(* IEC 61131-3 sources: STAR-PLC-Agent/results/raw/codex_matrix_resume_20261114/codex_deepseek/SELF011/functional/attempt_0001, 1 file *)

(* ---- test_program.st ---- *)
PROGRAM PLC_PRG
VAR
 BenchStep : UDINT := 0;
 BenchCalls : UDINT := 0;
 BenchDone : BOOL := FALSE;
 BenchUut0 : FB_Task;
 BenchUut1 : FB_Task;
 BenchUut2 : FB_Task;
 BenchUut3 : FB_Task;
 BenchUut4 : FB_Task;
 BenchUut5 : FB_Task;
 BenchUut6 : FB_Task;
 BenchUut7 : FB_Task;
 BenchUut8 : FB_Task;
 BenchUut9 : FB_Task;
 BenchUut10 : FB_Task;
 BenchUut11 : FB_Task;
 TraceIn_Start : ARRAY[0..147] OF BOOL;
 TraceIn_Stop : ARRAY[0..147] OF BOOL;
 TraceIn_Reset : ARRAY[0..147] OF BOOL;
 TraceIn_ExtendDone : ARRAY[0..147] OF BOOL;
 TraceIn_ClampDone : ARRAY[0..147] OF BOOL;
 TraceIn_ReleaseDone : ARRAY[0..147] OF BOOL;
 TraceIn_RetractDone : ARRAY[0..147] OF BOOL;
 TraceOut_Extend : ARRAY[0..147] OF BOOL;
 TraceOut_Clamp : ARRAY[0..147] OF BOOL;
 TraceOut_Release : ARRAY[0..147] OF BOOL;
 TraceOut_Retract : ARRAY[0..147] OF BOOL;
 TraceOut_Busy : ARRAY[0..147] OF BOOL;
 TraceOut_Done : ARRAY[0..147] OF BOOL;
END_VAR

IF NOT BenchDone THEN
 CASE BenchStep OF
 0:
   BenchUut0.Start := TRUE;
   BenchUut0.Stop := FALSE;
   BenchUut0.Reset := FALSE;
   BenchUut0.ExtendDone := FALSE;
   BenchUut0.ClampDone := FALSE;
   BenchUut0.ReleaseDone := FALSE;
   BenchUut0.RetractDone := FALSE;
   TraceIn_Start[0] := BenchUut0.Start;
   TraceIn_Stop[0] := BenchUut0.Stop;
   TraceIn_Reset[0] := BenchUut0.Reset;
   TraceIn_ExtendDone[0] := BenchUut0.ExtendDone;
   TraceIn_ClampDone[0] := BenchUut0.ClampDone;
   TraceIn_ReleaseDone[0] := BenchUut0.ReleaseDone;
   TraceIn_RetractDone[0] := BenchUut0.RetractDone;
   BenchUut0();
   TraceOut_Extend[0] := BenchUut0.Extend;
   TraceOut_Clamp[0] := BenchUut0.Clamp;
   TraceOut_Release[0] := BenchUut0.Release;
   TraceOut_Retract[0] := BenchUut0.Retract;
   TraceOut_Busy[0] := BenchUut0.Busy;
   TraceOut_Done[0] := BenchUut0.Done;
   BenchCalls := BenchCalls + 1;
 1:
   BenchUut0.Start := TRUE;
   BenchUut0.Stop := FALSE;
   BenchUut0.Reset := FALSE;
   BenchUut0.ExtendDone := FALSE;
   BenchUut0.ClampDone := FALSE;
   BenchUut0.ReleaseDone := FALSE;
   BenchUut0.RetractDone := TRUE;
   TraceIn_Start[1] := BenchUut0.Start;
   TraceIn_Stop[1] := BenchUut0.Stop;
   TraceIn_Reset[1] := BenchUut0.Reset;
   TraceIn_ExtendDone[1] := BenchUut0.ExtendDone;
   TraceIn_ClampDone[1] := BenchUut0.ClampDone;
   TraceIn_ReleaseDone[1] := BenchUut0.ReleaseDone;
   TraceIn_RetractDone[1] := BenchUut0.RetractDone;
   BenchUut0();
   TraceOut_Extend[1] := BenchUut0.Extend;
   TraceOut_Clamp[1] := BenchUut0.Clamp;
   TraceOut_Release[1] := BenchUut0.Release;
   TraceOut_Retract[1] := BenchUut0.Retract;
   TraceOut_Busy[1] := BenchUut0.Busy;
   TraceOut_Done[1] := BenchUut0.Done;
   BenchCalls := BenchCalls + 1;
 2:
   BenchUut0.Start := FALSE;
   BenchUut0.Stop := FALSE;
   BenchUut0.Reset := FALSE;
   BenchUut0.ExtendDone := FALSE;
   BenchUut0.ClampDone := FALSE;
   BenchUut0.ReleaseDone := FALSE;
   BenchUut0.RetractDone := FALSE;
   TraceIn_Start[2] := BenchUut0.Start;
   TraceIn_Stop[2] := BenchUut0.Stop;
   TraceIn_Reset[2] := BenchUut0.Reset;
   TraceIn_ExtendDone[2] := BenchUut0.ExtendDone;
   TraceIn_ClampDone[2] := BenchUut0.ClampDone;
   TraceIn_ReleaseDone[2] := BenchUut0.ReleaseDone;
   TraceIn_RetractDone[2] := BenchUut0.RetractDone;
   BenchUut0();
   TraceOut_Extend[2] := BenchUut0.Extend;
   TraceOut_Clamp[2] := BenchUut0.Clamp;
   TraceOut_Release[2] := BenchUut0.Release;
   TraceOut_Retract[2] := BenchUut0.Retract;
   TraceOut_Busy[2] := BenchUut0.Busy;
   TraceOut_Done[2] := BenchUut0.Done;
   BenchCalls := BenchCalls + 1;
 3:
   BenchUut0.Start := FALSE;
   BenchUut0.Stop := FALSE;
   BenchUut0.Reset := FALSE;
   BenchUut0.ExtendDone := TRUE;
   BenchUut0.ClampDone := FALSE;
   BenchUut0.ReleaseDone := FALSE;
   BenchUut0.RetractDone := FALSE;
   TraceIn_Start[3] := BenchUut0.Start;
   TraceIn_Stop[3] := BenchUut0.Stop;
   TraceIn_Reset[3] := BenchUut0.Reset;
   TraceIn_ExtendDone[3] := BenchUut0.ExtendDone;
   TraceIn_ClampDone[3] := BenchUut0.ClampDone;
   TraceIn_ReleaseDone[3] := BenchUut0.ReleaseDone;
   TraceIn_RetractDone[3] := BenchUut0.RetractDone;
   BenchUut0();
   TraceOut_Extend[3] := BenchUut0.Extend;
   TraceOut_Clamp[3] := BenchUut0.Clamp;
   TraceOut_Release[3] := BenchUut0.Release;
   TraceOut_Retract[3] := BenchUut0.Retract;
   TraceOut_Busy[3] := BenchUut0.Busy;
   TraceOut_Done[3] := BenchUut0.Done;
   BenchCalls := BenchCalls + 1;
 4:
   BenchUut0.Start := FALSE;
   BenchUut0.Stop := FALSE;
   BenchUut0.Reset := FALSE;
   BenchUut0.ExtendDone := FALSE;
   BenchUut0.ClampDone := TRUE;
   BenchUut0.ReleaseDone := FALSE;
   BenchUut0.RetractDone := FALSE;
   TraceIn_Start[4] := BenchUut0.Start;
   TraceIn_Stop[4] := BenchUut0.Stop;
   TraceIn_Reset[4] := BenchUut0.Reset;
   TraceIn_ExtendDone[4] := BenchUut0.ExtendDone;
   TraceIn_ClampDone[4] := BenchUut0.ClampDone;
   TraceIn_ReleaseDone[4] := BenchUut0.ReleaseDone;
   TraceIn_RetractDone[4] := BenchUut0.RetractDone;
   BenchUut0();
   TraceOut_Extend[4] := BenchUut0.Extend;
   TraceOut_Clamp[4] := BenchUut0.Clamp;
   TraceOut_Release[4] := BenchUut0.Release;
   TraceOut_Retract[4] := BenchUut0.Retract;
   TraceOut_Busy[4] := BenchUut0.Busy;
   TraceOut_Done[4] := BenchUut0.Done;
   BenchCalls := BenchCalls + 1;
 5:
   BenchUut0.Start := FALSE;
   BenchUut0.Stop := FALSE;
   BenchUut0.Reset := FALSE;
   BenchUut0.ExtendDone := FALSE;
   BenchUut0.ClampDone := FALSE;
   BenchUut0.ReleaseDone := TRUE;
   BenchUut0.RetractDone := FALSE;
   TraceIn_Start[5] := BenchUut0.Start;
   TraceIn_Stop[5] := BenchUut0.Stop;
   TraceIn_Reset[5] := BenchUut0.Reset;
   TraceIn_ExtendDone[5] := BenchUut0.ExtendDone;
   TraceIn_ClampDone[5] := BenchUut0.ClampDone;
   TraceIn_ReleaseDone[5] := BenchUut0.ReleaseDone;
   TraceIn_RetractDone[5] := BenchUut0.RetractDone;
   BenchUut0();
   TraceOut_Extend[5] := BenchUut0.Extend;
   TraceOut_Clamp[5] := BenchUut0.Clamp;
   TraceOut_Release[5] := BenchUut0.Release;
   TraceOut_Retract[5] := BenchUut0.Retract;
   TraceOut_Busy[5] := BenchUut0.Busy;
   TraceOut_Done[5] := BenchUut0.Done;
   BenchCalls := BenchCalls + 1;
 6:
   BenchUut0.Start := FALSE;
   BenchUut0.Stop := FALSE;
   BenchUut0.Reset := FALSE;
   BenchUut0.ExtendDone := FALSE;
   BenchUut0.ClampDone := FALSE;
   BenchUut0.ReleaseDone := FALSE;
   BenchUut0.RetractDone := TRUE;
   TraceIn_Start[6] := BenchUut0.Start;
   TraceIn_Stop[6] := BenchUut0.Stop;
   TraceIn_Reset[6] := BenchUut0.Reset;
   TraceIn_ExtendDone[6] := BenchUut0.ExtendDone;
   TraceIn_ClampDone[6] := BenchUut0.ClampDone;
   TraceIn_ReleaseDone[6] := BenchUut0.ReleaseDone;
   TraceIn_RetractDone[6] := BenchUut0.RetractDone;
   BenchUut0();
   TraceOut_Extend[6] := BenchUut0.Extend;
   TraceOut_Clamp[6] := BenchUut0.Clamp;
   TraceOut_Release[6] := BenchUut0.Release;
   TraceOut_Retract[6] := BenchUut0.Retract;
   TraceOut_Busy[6] := BenchUut0.Busy;
   TraceOut_Done[6] := BenchUut0.Done;
   BenchCalls := BenchCalls + 1;
 7:
   BenchUut0.Start := TRUE;
   BenchUut0.Stop := FALSE;
   BenchUut0.Reset := FALSE;
   BenchUut0.ExtendDone := FALSE;
   BenchUut0.ClampDone := FALSE;
   BenchUut0.ReleaseDone := FALSE;
   BenchUut0.RetractDone := FALSE;
   TraceIn_Start[7] := BenchUut0.Start;
   TraceIn_Stop[7] := BenchUut0.Stop;
   TraceIn_Reset[7] := BenchUut0.Reset;
   TraceIn_ExtendDone[7] := BenchUut0.ExtendDone;
   TraceIn_ClampDone[7] := BenchUut0.ClampDone;
   TraceIn_ReleaseDone[7] := BenchUut0.ReleaseDone;
   TraceIn_RetractDone[7] := BenchUut0.RetractDone;
   BenchUut0();
   TraceOut_Extend[7] := BenchUut0.Extend;
   TraceOut_Clamp[7] := BenchUut0.Clamp;
   TraceOut_Release[7] := BenchUut0.Release;
   TraceOut_Retract[7] := BenchUut0.Retract;
   TraceOut_Busy[7] := BenchUut0.Busy;
   TraceOut_Done[7] := BenchUut0.Done;
   BenchCalls := BenchCalls + 1;
 8:
   BenchUut0.Start := FALSE;
   BenchUut0.Stop := FALSE;
   BenchUut0.Reset := TRUE;
   BenchUut0.ExtendDone := FALSE;
   BenchUut0.ClampDone := FALSE;
   BenchUut0.ReleaseDone := FALSE;
   BenchUut0.RetractDone := FALSE;
   TraceIn_Start[8] := BenchUut0.Start;
   TraceIn_Stop[8] := BenchUut0.Stop;
   TraceIn_Reset[8] := BenchUut0.Reset;
   TraceIn_ExtendDone[8] := BenchUut0.ExtendDone;
   TraceIn_ClampDone[8] := BenchUut0.ClampDone;
   TraceIn_ReleaseDone[8] := BenchUut0.ReleaseDone;
   TraceIn_RetractDone[8] := BenchUut0.RetractDone;
   BenchUut0();
   TraceOut_Extend[8] := BenchUut0.Extend;
   TraceOut_Clamp[8] := BenchUut0.Clamp;
   TraceOut_Release[8] := BenchUut0.Release;
   TraceOut_Retract[8] := BenchUut0.Retract;
   TraceOut_Busy[8] := BenchUut0.Busy;
   TraceOut_Done[8] := BenchUut0.Done;
   BenchCalls := BenchCalls + 1;
 9:
   BenchUut1.Start := TRUE;
   BenchUut1.Stop := FALSE;
   BenchUut1.Reset := FALSE;
   BenchUut1.ExtendDone := TRUE;
   BenchUut1.ClampDone := TRUE;
   BenchUut1.ReleaseDone := TRUE;
   BenchUut1.RetractDone := TRUE;
   TraceIn_Start[9] := BenchUut1.Start;
   TraceIn_Stop[9] := BenchUut1.Stop;
   TraceIn_Reset[9] := BenchUut1.Reset;
   TraceIn_ExtendDone[9] := BenchUut1.ExtendDone;
   TraceIn_ClampDone[9] := BenchUut1.ClampDone;
   TraceIn_ReleaseDone[9] := BenchUut1.ReleaseDone;
   TraceIn_RetractDone[9] := BenchUut1.RetractDone;
   BenchUut1();
   TraceOut_Extend[9] := BenchUut1.Extend;
   TraceOut_Clamp[9] := BenchUut1.Clamp;
   TraceOut_Release[9] := BenchUut1.Release;
   TraceOut_Retract[9] := BenchUut1.Retract;
   TraceOut_Busy[9] := BenchUut1.Busy;
   TraceOut_Done[9] := BenchUut1.Done;
   BenchCalls := BenchCalls + 1;
 10:
   BenchUut1.Start := TRUE;
   BenchUut1.Stop := FALSE;
   BenchUut1.Reset := FALSE;
   BenchUut1.ExtendDone := TRUE;
   BenchUut1.ClampDone := TRUE;
   BenchUut1.ReleaseDone := TRUE;
   BenchUut1.RetractDone := TRUE;
   TraceIn_Start[10] := BenchUut1.Start;
   TraceIn_Stop[10] := BenchUut1.Stop;
   TraceIn_Reset[10] := BenchUut1.Reset;
   TraceIn_ExtendDone[10] := BenchUut1.ExtendDone;
   TraceIn_ClampDone[10] := BenchUut1.ClampDone;
   TraceIn_ReleaseDone[10] := BenchUut1.ReleaseDone;
   TraceIn_RetractDone[10] := BenchUut1.RetractDone;
   BenchUut1();
   TraceOut_Extend[10] := BenchUut1.Extend;
   TraceOut_Clamp[10] := BenchUut1.Clamp;
   TraceOut_Release[10] := BenchUut1.Release;
   TraceOut_Retract[10] := BenchUut1.Retract;
   TraceOut_Busy[10] := BenchUut1.Busy;
   TraceOut_Done[10] := BenchUut1.Done;
   BenchCalls := BenchCalls + 1;
 11:
   BenchUut1.Start := TRUE;
   BenchUut1.Stop := FALSE;
   BenchUut1.Reset := FALSE;
   BenchUut1.ExtendDone := TRUE;
   BenchUut1.ClampDone := TRUE;
   BenchUut1.ReleaseDone := TRUE;
   BenchUut1.RetractDone := TRUE;
   TraceIn_Start[11] := BenchUut1.Start;
   TraceIn_Stop[11] := BenchUut1.Stop;
   TraceIn_Reset[11] := BenchUut1.Reset;
   TraceIn_ExtendDone[11] := BenchUut1.ExtendDone;
   TraceIn_ClampDone[11] := BenchUut1.ClampDone;
   TraceIn_ReleaseDone[11] := BenchUut1.ReleaseDone;
   TraceIn_RetractDone[11] := BenchUut1.RetractDone;
   BenchUut1();
   TraceOut_Extend[11] := BenchUut1.Extend;
   TraceOut_Clamp[11] := BenchUut1.Clamp;
   TraceOut_Release[11] := BenchUut1.Release;
   TraceOut_Retract[11] := BenchUut1.Retract;
   TraceOut_Busy[11] := BenchUut1.Busy;
   TraceOut_Done[11] := BenchUut1.Done;
   BenchCalls := BenchCalls + 1;
 12:
   BenchUut1.Start := TRUE;
   BenchUut1.Stop := TRUE;
   BenchUut1.Reset := FALSE;
   BenchUut1.ExtendDone := TRUE;
   BenchUut1.ClampDone := TRUE;
   BenchUut1.ReleaseDone := TRUE;
   BenchUut1.RetractDone := TRUE;
   TraceIn_Start[12] := BenchUut1.Start;
   TraceIn_Stop[12] := BenchUut1.Stop;
   TraceIn_Reset[12] := BenchUut1.Reset;
   TraceIn_ExtendDone[12] := BenchUut1.ExtendDone;
   TraceIn_ClampDone[12] := BenchUut1.ClampDone;
   TraceIn_ReleaseDone[12] := BenchUut1.ReleaseDone;
   TraceIn_RetractDone[12] := BenchUut1.RetractDone;
   BenchUut1();
   TraceOut_Extend[12] := BenchUut1.Extend;
   TraceOut_Clamp[12] := BenchUut1.Clamp;
   TraceOut_Release[12] := BenchUut1.Release;
   TraceOut_Retract[12] := BenchUut1.Retract;
   TraceOut_Busy[12] := BenchUut1.Busy;
   TraceOut_Done[12] := BenchUut1.Done;
   BenchCalls := BenchCalls + 1;
 13:
   BenchUut1.Start := TRUE;
   BenchUut1.Stop := FALSE;
   BenchUut1.Reset := TRUE;
   BenchUut1.ExtendDone := TRUE;
   BenchUut1.ClampDone := TRUE;
   BenchUut1.ReleaseDone := TRUE;
   BenchUut1.RetractDone := TRUE;
   TraceIn_Start[13] := BenchUut1.Start;
   TraceIn_Stop[13] := BenchUut1.Stop;
   TraceIn_Reset[13] := BenchUut1.Reset;
   TraceIn_ExtendDone[13] := BenchUut1.ExtendDone;
   TraceIn_ClampDone[13] := BenchUut1.ClampDone;
   TraceIn_ReleaseDone[13] := BenchUut1.ReleaseDone;
   TraceIn_RetractDone[13] := BenchUut1.RetractDone;
   BenchUut1();
   TraceOut_Extend[13] := BenchUut1.Extend;
   TraceOut_Clamp[13] := BenchUut1.Clamp;
   TraceOut_Release[13] := BenchUut1.Release;
   TraceOut_Retract[13] := BenchUut1.Retract;
   TraceOut_Busy[13] := BenchUut1.Busy;
   TraceOut_Done[13] := BenchUut1.Done;
   BenchCalls := BenchCalls + 1;
 14:
   BenchUut2.Start := TRUE;
   BenchUut2.Stop := FALSE;
   BenchUut2.Reset := FALSE;
   BenchUut2.ExtendDone := FALSE;
   BenchUut2.ClampDone := FALSE;
   BenchUut2.ReleaseDone := FALSE;
   BenchUut2.RetractDone := TRUE;
   TraceIn_Start[14] := BenchUut2.Start;
   TraceIn_Stop[14] := BenchUut2.Stop;
   TraceIn_Reset[14] := BenchUut2.Reset;
   TraceIn_ExtendDone[14] := BenchUut2.ExtendDone;
   TraceIn_ClampDone[14] := BenchUut2.ClampDone;
   TraceIn_ReleaseDone[14] := BenchUut2.ReleaseDone;
   TraceIn_RetractDone[14] := BenchUut2.RetractDone;
   BenchUut2();
   TraceOut_Extend[14] := BenchUut2.Extend;
   TraceOut_Clamp[14] := BenchUut2.Clamp;
   TraceOut_Release[14] := BenchUut2.Release;
   TraceOut_Retract[14] := BenchUut2.Retract;
   TraceOut_Busy[14] := BenchUut2.Busy;
   TraceOut_Done[14] := BenchUut2.Done;
   BenchCalls := BenchCalls + 1;
 15:
   BenchUut2.Start := TRUE;
   BenchUut2.Stop := FALSE;
   BenchUut2.Reset := FALSE;
   BenchUut2.ExtendDone := TRUE;
   BenchUut2.ClampDone := FALSE;
   BenchUut2.ReleaseDone := FALSE;
   BenchUut2.RetractDone := FALSE;
   TraceIn_Start[15] := BenchUut2.Start;
   TraceIn_Stop[15] := BenchUut2.Stop;
   TraceIn_Reset[15] := BenchUut2.Reset;
   TraceIn_ExtendDone[15] := BenchUut2.ExtendDone;
   TraceIn_ClampDone[15] := BenchUut2.ClampDone;
   TraceIn_ReleaseDone[15] := BenchUut2.ReleaseDone;
   TraceIn_RetractDone[15] := BenchUut2.RetractDone;
   BenchUut2();
   TraceOut_Extend[15] := BenchUut2.Extend;
   TraceOut_Clamp[15] := BenchUut2.Clamp;
   TraceOut_Release[15] := BenchUut2.Release;
   TraceOut_Retract[15] := BenchUut2.Retract;
   TraceOut_Busy[15] := BenchUut2.Busy;
   TraceOut_Done[15] := BenchUut2.Done;
   BenchCalls := BenchCalls + 1;
 16:
   BenchUut2.Start := TRUE;
   BenchUut2.Stop := FALSE;
   BenchUut2.Reset := FALSE;
   BenchUut2.ExtendDone := FALSE;
   BenchUut2.ClampDone := FALSE;
   BenchUut2.ReleaseDone := FALSE;
   BenchUut2.RetractDone := FALSE;
   TraceIn_Start[16] := BenchUut2.Start;
   TraceIn_Stop[16] := BenchUut2.Stop;
   TraceIn_Reset[16] := BenchUut2.Reset;
   TraceIn_ExtendDone[16] := BenchUut2.ExtendDone;
   TraceIn_ClampDone[16] := BenchUut2.ClampDone;
   TraceIn_ReleaseDone[16] := BenchUut2.ReleaseDone;
   TraceIn_RetractDone[16] := BenchUut2.RetractDone;
   BenchUut2();
   TraceOut_Extend[16] := BenchUut2.Extend;
   TraceOut_Clamp[16] := BenchUut2.Clamp;
   TraceOut_Release[16] := BenchUut2.Release;
   TraceOut_Retract[16] := BenchUut2.Retract;
   TraceOut_Busy[16] := BenchUut2.Busy;
   TraceOut_Done[16] := BenchUut2.Done;
   BenchCalls := BenchCalls + 1;
 17:
   BenchUut2.Start := FALSE;
   BenchUut2.Stop := FALSE;
   BenchUut2.Reset := FALSE;
   BenchUut2.ExtendDone := FALSE;
   BenchUut2.ClampDone := TRUE;
   BenchUut2.ReleaseDone := FALSE;
   BenchUut2.RetractDone := FALSE;
   TraceIn_Start[17] := BenchUut2.Start;
   TraceIn_Stop[17] := BenchUut2.Stop;
   TraceIn_Reset[17] := BenchUut2.Reset;
   TraceIn_ExtendDone[17] := BenchUut2.ExtendDone;
   TraceIn_ClampDone[17] := BenchUut2.ClampDone;
   TraceIn_ReleaseDone[17] := BenchUut2.ReleaseDone;
   TraceIn_RetractDone[17] := BenchUut2.RetractDone;
   BenchUut2();
   TraceOut_Extend[17] := BenchUut2.Extend;
   TraceOut_Clamp[17] := BenchUut2.Clamp;
   TraceOut_Release[17] := BenchUut2.Release;
   TraceOut_Retract[17] := BenchUut2.Retract;
   TraceOut_Busy[17] := BenchUut2.Busy;
   TraceOut_Done[17] := BenchUut2.Done;
   BenchCalls := BenchCalls + 1;
 18:
   BenchUut2.Start := FALSE;
   BenchUut2.Stop := FALSE;
   BenchUut2.Reset := FALSE;
   BenchUut2.ExtendDone := FALSE;
   BenchUut2.ClampDone := FALSE;
   BenchUut2.ReleaseDone := FALSE;
   BenchUut2.RetractDone := FALSE;
   TraceIn_Start[18] := BenchUut2.Start;
   TraceIn_Stop[18] := BenchUut2.Stop;
   TraceIn_Reset[18] := BenchUut2.Reset;
   TraceIn_ExtendDone[18] := BenchUut2.ExtendDone;
   TraceIn_ClampDone[18] := BenchUut2.ClampDone;
   TraceIn_ReleaseDone[18] := BenchUut2.ReleaseDone;
   TraceIn_RetractDone[18] := BenchUut2.RetractDone;
   BenchUut2();
   TraceOut_Extend[18] := BenchUut2.Extend;
   TraceOut_Clamp[18] := BenchUut2.Clamp;
   TraceOut_Release[18] := BenchUut2.Release;
   TraceOut_Retract[18] := BenchUut2.Retract;
   TraceOut_Busy[18] := BenchUut2.Busy;
   TraceOut_Done[18] := BenchUut2.Done;
   BenchCalls := BenchCalls + 1;
 19:
   BenchUut2.Start := FALSE;
   BenchUut2.Stop := FALSE;
   BenchUut2.Reset := FALSE;
   BenchUut2.ExtendDone := FALSE;
   BenchUut2.ClampDone := FALSE;
   BenchUut2.ReleaseDone := TRUE;
   BenchUut2.RetractDone := FALSE;
   TraceIn_Start[19] := BenchUut2.Start;
   TraceIn_Stop[19] := BenchUut2.Stop;
   TraceIn_Reset[19] := BenchUut2.Reset;
   TraceIn_ExtendDone[19] := BenchUut2.ExtendDone;
   TraceIn_ClampDone[19] := BenchUut2.ClampDone;
   TraceIn_ReleaseDone[19] := BenchUut2.ReleaseDone;
   TraceIn_RetractDone[19] := BenchUut2.RetractDone;
   BenchUut2();
   TraceOut_Extend[19] := BenchUut2.Extend;
   TraceOut_Clamp[19] := BenchUut2.Clamp;
   TraceOut_Release[19] := BenchUut2.Release;
   TraceOut_Retract[19] := BenchUut2.Retract;
   TraceOut_Busy[19] := BenchUut2.Busy;
   TraceOut_Done[19] := BenchUut2.Done;
   BenchCalls := BenchCalls + 1;
 20:
   BenchUut2.Start := FALSE;
   BenchUut2.Stop := FALSE;
   BenchUut2.Reset := FALSE;
   BenchUut2.ExtendDone := FALSE;
   BenchUut2.ClampDone := FALSE;
   BenchUut2.ReleaseDone := FALSE;
   BenchUut2.RetractDone := FALSE;
   TraceIn_Start[20] := BenchUut2.Start;
   TraceIn_Stop[20] := BenchUut2.Stop;
   TraceIn_Reset[20] := BenchUut2.Reset;
   TraceIn_ExtendDone[20] := BenchUut2.ExtendDone;
   TraceIn_ClampDone[20] := BenchUut2.ClampDone;
   TraceIn_ReleaseDone[20] := BenchUut2.ReleaseDone;
   TraceIn_RetractDone[20] := BenchUut2.RetractDone;
   BenchUut2();
   TraceOut_Extend[20] := BenchUut2.Extend;
   TraceOut_Clamp[20] := BenchUut2.Clamp;
   TraceOut_Release[20] := BenchUut2.Release;
   TraceOut_Retract[20] := BenchUut2.Retract;
   TraceOut_Busy[20] := BenchUut2.Busy;
   TraceOut_Done[20] := BenchUut2.Done;
   BenchCalls := BenchCalls + 1;
 21:
   BenchUut2.Start := FALSE;
   BenchUut2.Stop := FALSE;
   BenchUut2.Reset := FALSE;
   BenchUut2.ExtendDone := FALSE;
   BenchUut2.ClampDone := FALSE;
   BenchUut2.ReleaseDone := FALSE;
   BenchUut2.RetractDone := TRUE;
   TraceIn_Start[21] := BenchUut2.Start;
   TraceIn_Stop[21] := BenchUut2.Stop;
   TraceIn_Reset[21] := BenchUut2.Reset;
   TraceIn_ExtendDone[21] := BenchUut2.ExtendDone;
   TraceIn_ClampDone[21] := BenchUut2.ClampDone;
   TraceIn_ReleaseDone[21] := BenchUut2.ReleaseDone;
   TraceIn_RetractDone[21] := BenchUut2.RetractDone;
   BenchUut2();
   TraceOut_Extend[21] := BenchUut2.Extend;
   TraceOut_Clamp[21] := BenchUut2.Clamp;
   TraceOut_Release[21] := BenchUut2.Release;
   TraceOut_Retract[21] := BenchUut2.Retract;
   TraceOut_Busy[21] := BenchUut2.Busy;
   TraceOut_Done[21] := BenchUut2.Done;
   BenchCalls := BenchCalls + 1;
 22:
   BenchUut2.Start := FALSE;
   BenchUut2.Stop := TRUE;
   BenchUut2.Reset := FALSE;
   BenchUut2.ExtendDone := FALSE;
   BenchUut2.ClampDone := FALSE;
   BenchUut2.ReleaseDone := FALSE;
   BenchUut2.RetractDone := TRUE;
   TraceIn_Start[22] := BenchUut2.Start;
   TraceIn_Stop[22] := BenchUut2.Stop;
   TraceIn_Reset[22] := BenchUut2.Reset;
   TraceIn_ExtendDone[22] := BenchUut2.ExtendDone;
   TraceIn_ClampDone[22] := BenchUut2.ClampDone;
   TraceIn_ReleaseDone[22] := BenchUut2.ReleaseDone;
   TraceIn_RetractDone[22] := BenchUut2.RetractDone;
   BenchUut2();
   TraceOut_Extend[22] := BenchUut2.Extend;
   TraceOut_Clamp[22] := BenchUut2.Clamp;
   TraceOut_Release[22] := BenchUut2.Release;
   TraceOut_Retract[22] := BenchUut2.Retract;
   TraceOut_Busy[22] := BenchUut2.Busy;
   TraceOut_Done[22] := BenchUut2.Done;
   BenchCalls := BenchCalls + 1;
 23:
   BenchUut2.Start := TRUE;
   BenchUut2.Stop := FALSE;
   BenchUut2.Reset := FALSE;
   BenchUut2.ExtendDone := FALSE;
   BenchUut2.ClampDone := FALSE;
   BenchUut2.ReleaseDone := FALSE;
   BenchUut2.RetractDone := TRUE;
   TraceIn_Start[23] := BenchUut2.Start;
   TraceIn_Stop[23] := BenchUut2.Stop;
   TraceIn_Reset[23] := BenchUut2.Reset;
   TraceIn_ExtendDone[23] := BenchUut2.ExtendDone;
   TraceIn_ClampDone[23] := BenchUut2.ClampDone;
   TraceIn_ReleaseDone[23] := BenchUut2.ReleaseDone;
   TraceIn_RetractDone[23] := BenchUut2.RetractDone;
   BenchUut2();
   TraceOut_Extend[23] := BenchUut2.Extend;
   TraceOut_Clamp[23] := BenchUut2.Clamp;
   TraceOut_Release[23] := BenchUut2.Release;
   TraceOut_Retract[23] := BenchUut2.Retract;
   TraceOut_Busy[23] := BenchUut2.Busy;
   TraceOut_Done[23] := BenchUut2.Done;
   BenchCalls := BenchCalls + 1;
 24:
   BenchUut3.Start := TRUE;
   BenchUut3.Stop := FALSE;
   BenchUut3.Reset := FALSE;
   BenchUut3.ExtendDone := FALSE;
   BenchUut3.ClampDone := FALSE;
   BenchUut3.ReleaseDone := FALSE;
   BenchUut3.RetractDone := FALSE;
   TraceIn_Start[24] := BenchUut3.Start;
   TraceIn_Stop[24] := BenchUut3.Stop;
   TraceIn_Reset[24] := BenchUut3.Reset;
   TraceIn_ExtendDone[24] := BenchUut3.ExtendDone;
   TraceIn_ClampDone[24] := BenchUut3.ClampDone;
   TraceIn_ReleaseDone[24] := BenchUut3.ReleaseDone;
   TraceIn_RetractDone[24] := BenchUut3.RetractDone;
   BenchUut3();
   TraceOut_Extend[24] := BenchUut3.Extend;
   TraceOut_Clamp[24] := BenchUut3.Clamp;
   TraceOut_Release[24] := BenchUut3.Release;
   TraceOut_Retract[24] := BenchUut3.Retract;
   TraceOut_Busy[24] := BenchUut3.Busy;
   TraceOut_Done[24] := BenchUut3.Done;
   BenchCalls := BenchCalls + 1;
 25:
   BenchUut3.Start := TRUE;
   BenchUut3.Stop := FALSE;
   BenchUut3.Reset := FALSE;
   BenchUut3.ExtendDone := FALSE;
   BenchUut3.ClampDone := FALSE;
   BenchUut3.ReleaseDone := FALSE;
   BenchUut3.RetractDone := TRUE;
   TraceIn_Start[25] := BenchUut3.Start;
   TraceIn_Stop[25] := BenchUut3.Stop;
   TraceIn_Reset[25] := BenchUut3.Reset;
   TraceIn_ExtendDone[25] := BenchUut3.ExtendDone;
   TraceIn_ClampDone[25] := BenchUut3.ClampDone;
   TraceIn_ReleaseDone[25] := BenchUut3.ReleaseDone;
   TraceIn_RetractDone[25] := BenchUut3.RetractDone;
   BenchUut3();
   TraceOut_Extend[25] := BenchUut3.Extend;
   TraceOut_Clamp[25] := BenchUut3.Clamp;
   TraceOut_Release[25] := BenchUut3.Release;
   TraceOut_Retract[25] := BenchUut3.Retract;
   TraceOut_Busy[25] := BenchUut3.Busy;
   TraceOut_Done[25] := BenchUut3.Done;
   BenchCalls := BenchCalls + 1;
 26:
   BenchUut3.Start := FALSE;
   BenchUut3.Stop := FALSE;
   BenchUut3.Reset := FALSE;
   BenchUut3.ExtendDone := FALSE;
   BenchUut3.ClampDone := FALSE;
   BenchUut3.ReleaseDone := FALSE;
   BenchUut3.RetractDone := FALSE;
   TraceIn_Start[26] := BenchUut3.Start;
   TraceIn_Stop[26] := BenchUut3.Stop;
   TraceIn_Reset[26] := BenchUut3.Reset;
   TraceIn_ExtendDone[26] := BenchUut3.ExtendDone;
   TraceIn_ClampDone[26] := BenchUut3.ClampDone;
   TraceIn_ReleaseDone[26] := BenchUut3.ReleaseDone;
   TraceIn_RetractDone[26] := BenchUut3.RetractDone;
   BenchUut3();
   TraceOut_Extend[26] := BenchUut3.Extend;
   TraceOut_Clamp[26] := BenchUut3.Clamp;
   TraceOut_Release[26] := BenchUut3.Release;
   TraceOut_Retract[26] := BenchUut3.Retract;
   TraceOut_Busy[26] := BenchUut3.Busy;
   TraceOut_Done[26] := BenchUut3.Done;
   BenchCalls := BenchCalls + 1;
 27:
   BenchUut3.Start := FALSE;
   BenchUut3.Stop := FALSE;
   BenchUut3.Reset := FALSE;
   BenchUut3.ExtendDone := TRUE;
   BenchUut3.ClampDone := FALSE;
   BenchUut3.ReleaseDone := FALSE;
   BenchUut3.RetractDone := FALSE;
   TraceIn_Start[27] := BenchUut3.Start;
   TraceIn_Stop[27] := BenchUut3.Stop;
   TraceIn_Reset[27] := BenchUut3.Reset;
   TraceIn_ExtendDone[27] := BenchUut3.ExtendDone;
   TraceIn_ClampDone[27] := BenchUut3.ClampDone;
   TraceIn_ReleaseDone[27] := BenchUut3.ReleaseDone;
   TraceIn_RetractDone[27] := BenchUut3.RetractDone;
   BenchUut3();
   TraceOut_Extend[27] := BenchUut3.Extend;
   TraceOut_Clamp[27] := BenchUut3.Clamp;
   TraceOut_Release[27] := BenchUut3.Release;
   TraceOut_Retract[27] := BenchUut3.Retract;
   TraceOut_Busy[27] := BenchUut3.Busy;
   TraceOut_Done[27] := BenchUut3.Done;
   BenchCalls := BenchCalls + 1;
 28:
   BenchUut3.Start := FALSE;
   BenchUut3.Stop := FALSE;
   BenchUut3.Reset := FALSE;
   BenchUut3.ExtendDone := FALSE;
   BenchUut3.ClampDone := FALSE;
   BenchUut3.ReleaseDone := FALSE;
   BenchUut3.RetractDone := FALSE;
   TraceIn_Start[28] := BenchUut3.Start;
   TraceIn_Stop[28] := BenchUut3.Stop;
   TraceIn_Reset[28] := BenchUut3.Reset;
   TraceIn_ExtendDone[28] := BenchUut3.ExtendDone;
   TraceIn_ClampDone[28] := BenchUut3.ClampDone;
   TraceIn_ReleaseDone[28] := BenchUut3.ReleaseDone;
   TraceIn_RetractDone[28] := BenchUut3.RetractDone;
   BenchUut3();
   TraceOut_Extend[28] := BenchUut3.Extend;
   TraceOut_Clamp[28] := BenchUut3.Clamp;
   TraceOut_Release[28] := BenchUut3.Release;
   TraceOut_Retract[28] := BenchUut3.Retract;
   TraceOut_Busy[28] := BenchUut3.Busy;
   TraceOut_Done[28] := BenchUut3.Done;
   BenchCalls := BenchCalls + 1;
 29:
   BenchUut4.Start := FALSE;
   BenchUut4.Stop := FALSE;
   BenchUut4.Reset := TRUE;
   BenchUut4.ExtendDone := FALSE;
   BenchUut4.ClampDone := FALSE;
   BenchUut4.ReleaseDone := FALSE;
   BenchUut4.RetractDone := TRUE;
   TraceIn_Start[29] := BenchUut4.Start;
   TraceIn_Stop[29] := BenchUut4.Stop;
   TraceIn_Reset[29] := BenchUut4.Reset;
   TraceIn_ExtendDone[29] := BenchUut4.ExtendDone;
   TraceIn_ClampDone[29] := BenchUut4.ClampDone;
   TraceIn_ReleaseDone[29] := BenchUut4.ReleaseDone;
   TraceIn_RetractDone[29] := BenchUut4.RetractDone;
   BenchUut4();
   TraceOut_Extend[29] := BenchUut4.Extend;
   TraceOut_Clamp[29] := BenchUut4.Clamp;
   TraceOut_Release[29] := BenchUut4.Release;
   TraceOut_Retract[29] := BenchUut4.Retract;
   TraceOut_Busy[29] := BenchUut4.Busy;
   TraceOut_Done[29] := BenchUut4.Done;
   BenchCalls := BenchCalls + 1;
 30:
   BenchUut4.Start := FALSE;
   BenchUut4.Stop := FALSE;
   BenchUut4.Reset := FALSE;
   BenchUut4.ExtendDone := FALSE;
   BenchUut4.ClampDone := FALSE;
   BenchUut4.ReleaseDone := FALSE;
   BenchUut4.RetractDone := TRUE;
   TraceIn_Start[30] := BenchUut4.Start;
   TraceIn_Stop[30] := BenchUut4.Stop;
   TraceIn_Reset[30] := BenchUut4.Reset;
   TraceIn_ExtendDone[30] := BenchUut4.ExtendDone;
   TraceIn_ClampDone[30] := BenchUut4.ClampDone;
   TraceIn_ReleaseDone[30] := BenchUut4.ReleaseDone;
   TraceIn_RetractDone[30] := BenchUut4.RetractDone;
   BenchUut4();
   TraceOut_Extend[30] := BenchUut4.Extend;
   TraceOut_Clamp[30] := BenchUut4.Clamp;
   TraceOut_Release[30] := BenchUut4.Release;
   TraceOut_Retract[30] := BenchUut4.Retract;
   TraceOut_Busy[30] := BenchUut4.Busy;
   TraceOut_Done[30] := BenchUut4.Done;
   BenchCalls := BenchCalls + 1;
 31:
   BenchUut4.Start := TRUE;
   BenchUut4.Stop := FALSE;
   BenchUut4.Reset := FALSE;
   BenchUut4.ExtendDone := FALSE;
   BenchUut4.ClampDone := FALSE;
   BenchUut4.ReleaseDone := FALSE;
   BenchUut4.RetractDone := TRUE;
   TraceIn_Start[31] := BenchUut4.Start;
   TraceIn_Stop[31] := BenchUut4.Stop;
   TraceIn_Reset[31] := BenchUut4.Reset;
   TraceIn_ExtendDone[31] := BenchUut4.ExtendDone;
   TraceIn_ClampDone[31] := BenchUut4.ClampDone;
   TraceIn_ReleaseDone[31] := BenchUut4.ReleaseDone;
   TraceIn_RetractDone[31] := BenchUut4.RetractDone;
   BenchUut4();
   TraceOut_Extend[31] := BenchUut4.Extend;
   TraceOut_Clamp[31] := BenchUut4.Clamp;
   TraceOut_Release[31] := BenchUut4.Release;
   TraceOut_Retract[31] := BenchUut4.Retract;
   TraceOut_Busy[31] := BenchUut4.Busy;
   TraceOut_Done[31] := BenchUut4.Done;
   BenchCalls := BenchCalls + 1;
 32:
   BenchUut4.Start := FALSE;
   BenchUut4.Stop := FALSE;
   BenchUut4.Reset := FALSE;
   BenchUut4.ExtendDone := FALSE;
   BenchUut4.ClampDone := FALSE;
   BenchUut4.ReleaseDone := FALSE;
   BenchUut4.RetractDone := FALSE;
   TraceIn_Start[32] := BenchUut4.Start;
   TraceIn_Stop[32] := BenchUut4.Stop;
   TraceIn_Reset[32] := BenchUut4.Reset;
   TraceIn_ExtendDone[32] := BenchUut4.ExtendDone;
   TraceIn_ClampDone[32] := BenchUut4.ClampDone;
   TraceIn_ReleaseDone[32] := BenchUut4.ReleaseDone;
   TraceIn_RetractDone[32] := BenchUut4.RetractDone;
   BenchUut4();
   TraceOut_Extend[32] := BenchUut4.Extend;
   TraceOut_Clamp[32] := BenchUut4.Clamp;
   TraceOut_Release[32] := BenchUut4.Release;
   TraceOut_Retract[32] := BenchUut4.Retract;
   TraceOut_Busy[32] := BenchUut4.Busy;
   TraceOut_Done[32] := BenchUut4.Done;
   BenchCalls := BenchCalls + 1;
 33:
   BenchUut4.Start := FALSE;
   BenchUut4.Stop := FALSE;
   BenchUut4.Reset := FALSE;
   BenchUut4.ExtendDone := FALSE;
   BenchUut4.ClampDone := FALSE;
   BenchUut4.ReleaseDone := FALSE;
   BenchUut4.RetractDone := FALSE;
   TraceIn_Start[33] := BenchUut4.Start;
   TraceIn_Stop[33] := BenchUut4.Stop;
   TraceIn_Reset[33] := BenchUut4.Reset;
   TraceIn_ExtendDone[33] := BenchUut4.ExtendDone;
   TraceIn_ClampDone[33] := BenchUut4.ClampDone;
   TraceIn_ReleaseDone[33] := BenchUut4.ReleaseDone;
   TraceIn_RetractDone[33] := BenchUut4.RetractDone;
   BenchUut4();
   TraceOut_Extend[33] := BenchUut4.Extend;
   TraceOut_Clamp[33] := BenchUut4.Clamp;
   TraceOut_Release[33] := BenchUut4.Release;
   TraceOut_Retract[33] := BenchUut4.Retract;
   TraceOut_Busy[33] := BenchUut4.Busy;
   TraceOut_Done[33] := BenchUut4.Done;
   BenchCalls := BenchCalls + 1;
 34:
   BenchUut4.Start := FALSE;
   BenchUut4.Stop := FALSE;
   BenchUut4.Reset := FALSE;
   BenchUut4.ExtendDone := TRUE;
   BenchUut4.ClampDone := FALSE;
   BenchUut4.ReleaseDone := FALSE;
   BenchUut4.RetractDone := FALSE;
   TraceIn_Start[34] := BenchUut4.Start;
   TraceIn_Stop[34] := BenchUut4.Stop;
   TraceIn_Reset[34] := BenchUut4.Reset;
   TraceIn_ExtendDone[34] := BenchUut4.ExtendDone;
   TraceIn_ClampDone[34] := BenchUut4.ClampDone;
   TraceIn_ReleaseDone[34] := BenchUut4.ReleaseDone;
   TraceIn_RetractDone[34] := BenchUut4.RetractDone;
   BenchUut4();
   TraceOut_Extend[34] := BenchUut4.Extend;
   TraceOut_Clamp[34] := BenchUut4.Clamp;
   TraceOut_Release[34] := BenchUut4.Release;
   TraceOut_Retract[34] := BenchUut4.Retract;
   TraceOut_Busy[34] := BenchUut4.Busy;
   TraceOut_Done[34] := BenchUut4.Done;
   BenchCalls := BenchCalls + 1;
 35:
   BenchUut4.Start := FALSE;
   BenchUut4.Stop := FALSE;
   BenchUut4.Reset := FALSE;
   BenchUut4.ExtendDone := FALSE;
   BenchUut4.ClampDone := FALSE;
   BenchUut4.ReleaseDone := FALSE;
   BenchUut4.RetractDone := FALSE;
   TraceIn_Start[35] := BenchUut4.Start;
   TraceIn_Stop[35] := BenchUut4.Stop;
   TraceIn_Reset[35] := BenchUut4.Reset;
   TraceIn_ExtendDone[35] := BenchUut4.ExtendDone;
   TraceIn_ClampDone[35] := BenchUut4.ClampDone;
   TraceIn_ReleaseDone[35] := BenchUut4.ReleaseDone;
   TraceIn_RetractDone[35] := BenchUut4.RetractDone;
   BenchUut4();
   TraceOut_Extend[35] := BenchUut4.Extend;
   TraceOut_Clamp[35] := BenchUut4.Clamp;
   TraceOut_Release[35] := BenchUut4.Release;
   TraceOut_Retract[35] := BenchUut4.Retract;
   TraceOut_Busy[35] := BenchUut4.Busy;
   TraceOut_Done[35] := BenchUut4.Done;
   BenchCalls := BenchCalls + 1;
 36:
   BenchUut4.Start := FALSE;
   BenchUut4.Stop := FALSE;
   BenchUut4.Reset := FALSE;
   BenchUut4.ExtendDone := FALSE;
   BenchUut4.ClampDone := FALSE;
   BenchUut4.ReleaseDone := FALSE;
   BenchUut4.RetractDone := FALSE;
   TraceIn_Start[36] := BenchUut4.Start;
   TraceIn_Stop[36] := BenchUut4.Stop;
   TraceIn_Reset[36] := BenchUut4.Reset;
   TraceIn_ExtendDone[36] := BenchUut4.ExtendDone;
   TraceIn_ClampDone[36] := BenchUut4.ClampDone;
   TraceIn_ReleaseDone[36] := BenchUut4.ReleaseDone;
   TraceIn_RetractDone[36] := BenchUut4.RetractDone;
   BenchUut4();
   TraceOut_Extend[36] := BenchUut4.Extend;
   TraceOut_Clamp[36] := BenchUut4.Clamp;
   TraceOut_Release[36] := BenchUut4.Release;
   TraceOut_Retract[36] := BenchUut4.Retract;
   TraceOut_Busy[36] := BenchUut4.Busy;
   TraceOut_Done[36] := BenchUut4.Done;
   BenchCalls := BenchCalls + 1;
 37:
   BenchUut4.Start := FALSE;
   BenchUut4.Stop := FALSE;
   BenchUut4.Reset := FALSE;
   BenchUut4.ExtendDone := FALSE;
   BenchUut4.ClampDone := FALSE;
   BenchUut4.ReleaseDone := FALSE;
   BenchUut4.RetractDone := FALSE;
   TraceIn_Start[37] := BenchUut4.Start;
   TraceIn_Stop[37] := BenchUut4.Stop;
   TraceIn_Reset[37] := BenchUut4.Reset;
   TraceIn_ExtendDone[37] := BenchUut4.ExtendDone;
   TraceIn_ClampDone[37] := BenchUut4.ClampDone;
   TraceIn_ReleaseDone[37] := BenchUut4.ReleaseDone;
   TraceIn_RetractDone[37] := BenchUut4.RetractDone;
   BenchUut4();
   TraceOut_Extend[37] := BenchUut4.Extend;
   TraceOut_Clamp[37] := BenchUut4.Clamp;
   TraceOut_Release[37] := BenchUut4.Release;
   TraceOut_Retract[37] := BenchUut4.Retract;
   TraceOut_Busy[37] := BenchUut4.Busy;
   TraceOut_Done[37] := BenchUut4.Done;
   BenchCalls := BenchCalls + 1;
 38:
   BenchUut4.Start := FALSE;
   BenchUut4.Stop := FALSE;
   BenchUut4.Reset := FALSE;
   BenchUut4.ExtendDone := FALSE;
   BenchUut4.ClampDone := TRUE;
   BenchUut4.ReleaseDone := FALSE;
   BenchUut4.RetractDone := FALSE;
   TraceIn_Start[38] := BenchUut4.Start;
   TraceIn_Stop[38] := BenchUut4.Stop;
   TraceIn_Reset[38] := BenchUut4.Reset;
   TraceIn_ExtendDone[38] := BenchUut4.ExtendDone;
   TraceIn_ClampDone[38] := BenchUut4.ClampDone;
   TraceIn_ReleaseDone[38] := BenchUut4.ReleaseDone;
   TraceIn_RetractDone[38] := BenchUut4.RetractDone;
   BenchUut4();
   TraceOut_Extend[38] := BenchUut4.Extend;
   TraceOut_Clamp[38] := BenchUut4.Clamp;
   TraceOut_Release[38] := BenchUut4.Release;
   TraceOut_Retract[38] := BenchUut4.Retract;
   TraceOut_Busy[38] := BenchUut4.Busy;
   TraceOut_Done[38] := BenchUut4.Done;
   BenchCalls := BenchCalls + 1;
 39:
   BenchUut4.Start := FALSE;
   BenchUut4.Stop := FALSE;
   BenchUut4.Reset := FALSE;
   BenchUut4.ExtendDone := FALSE;
   BenchUut4.ClampDone := FALSE;
   BenchUut4.ReleaseDone := FALSE;
   BenchUut4.RetractDone := FALSE;
   TraceIn_Start[39] := BenchUut4.Start;
   TraceIn_Stop[39] := BenchUut4.Stop;
   TraceIn_Reset[39] := BenchUut4.Reset;
   TraceIn_ExtendDone[39] := BenchUut4.ExtendDone;
   TraceIn_ClampDone[39] := BenchUut4.ClampDone;
   TraceIn_ReleaseDone[39] := BenchUut4.ReleaseDone;
   TraceIn_RetractDone[39] := BenchUut4.RetractDone;
   BenchUut4();
   TraceOut_Extend[39] := BenchUut4.Extend;
   TraceOut_Clamp[39] := BenchUut4.Clamp;
   TraceOut_Release[39] := BenchUut4.Release;
   TraceOut_Retract[39] := BenchUut4.Retract;
   TraceOut_Busy[39] := BenchUut4.Busy;
   TraceOut_Done[39] := BenchUut4.Done;
   BenchCalls := BenchCalls + 1;
 40:
   BenchUut4.Start := FALSE;
   BenchUut4.Stop := FALSE;
   BenchUut4.Reset := FALSE;
   BenchUut4.ExtendDone := FALSE;
   BenchUut4.ClampDone := FALSE;
   BenchUut4.ReleaseDone := FALSE;
   BenchUut4.RetractDone := FALSE;
   TraceIn_Start[40] := BenchUut4.Start;
   TraceIn_Stop[40] := BenchUut4.Stop;
   TraceIn_Reset[40] := BenchUut4.Reset;
   TraceIn_ExtendDone[40] := BenchUut4.ExtendDone;
   TraceIn_ClampDone[40] := BenchUut4.ClampDone;
   TraceIn_ReleaseDone[40] := BenchUut4.ReleaseDone;
   TraceIn_RetractDone[40] := BenchUut4.RetractDone;
   BenchUut4();
   TraceOut_Extend[40] := BenchUut4.Extend;
   TraceOut_Clamp[40] := BenchUut4.Clamp;
   TraceOut_Release[40] := BenchUut4.Release;
   TraceOut_Retract[40] := BenchUut4.Retract;
   TraceOut_Busy[40] := BenchUut4.Busy;
   TraceOut_Done[40] := BenchUut4.Done;
   BenchCalls := BenchCalls + 1;
 41:
   BenchUut4.Start := FALSE;
   BenchUut4.Stop := FALSE;
   BenchUut4.Reset := FALSE;
   BenchUut4.ExtendDone := FALSE;
   BenchUut4.ClampDone := FALSE;
   BenchUut4.ReleaseDone := FALSE;
   BenchUut4.RetractDone := FALSE;
   TraceIn_Start[41] := BenchUut4.Start;
   TraceIn_Stop[41] := BenchUut4.Stop;
   TraceIn_Reset[41] := BenchUut4.Reset;
   TraceIn_ExtendDone[41] := BenchUut4.ExtendDone;
   TraceIn_ClampDone[41] := BenchUut4.ClampDone;
   TraceIn_ReleaseDone[41] := BenchUut4.ReleaseDone;
   TraceIn_RetractDone[41] := BenchUut4.RetractDone;
   BenchUut4();
   TraceOut_Extend[41] := BenchUut4.Extend;
   TraceOut_Clamp[41] := BenchUut4.Clamp;
   TraceOut_Release[41] := BenchUut4.Release;
   TraceOut_Retract[41] := BenchUut4.Retract;
   TraceOut_Busy[41] := BenchUut4.Busy;
   TraceOut_Done[41] := BenchUut4.Done;
   BenchCalls := BenchCalls + 1;
 42:
   BenchUut4.Start := FALSE;
   BenchUut4.Stop := FALSE;
   BenchUut4.Reset := FALSE;
   BenchUut4.ExtendDone := FALSE;
   BenchUut4.ClampDone := FALSE;
   BenchUut4.ReleaseDone := TRUE;
   BenchUut4.RetractDone := FALSE;
   TraceIn_Start[42] := BenchUut4.Start;
   TraceIn_Stop[42] := BenchUut4.Stop;
   TraceIn_Reset[42] := BenchUut4.Reset;
   TraceIn_ExtendDone[42] := BenchUut4.ExtendDone;
   TraceIn_ClampDone[42] := BenchUut4.ClampDone;
   TraceIn_ReleaseDone[42] := BenchUut4.ReleaseDone;
   TraceIn_RetractDone[42] := BenchUut4.RetractDone;
   BenchUut4();
   TraceOut_Extend[42] := BenchUut4.Extend;
   TraceOut_Clamp[42] := BenchUut4.Clamp;
   TraceOut_Release[42] := BenchUut4.Release;
   TraceOut_Retract[42] := BenchUut4.Retract;
   TraceOut_Busy[42] := BenchUut4.Busy;
   TraceOut_Done[42] := BenchUut4.Done;
   BenchCalls := BenchCalls + 1;
 43:
   BenchUut4.Start := FALSE;
   BenchUut4.Stop := FALSE;
   BenchUut4.Reset := FALSE;
   BenchUut4.ExtendDone := FALSE;
   BenchUut4.ClampDone := FALSE;
   BenchUut4.ReleaseDone := FALSE;
   BenchUut4.RetractDone := FALSE;
   TraceIn_Start[43] := BenchUut4.Start;
   TraceIn_Stop[43] := BenchUut4.Stop;
   TraceIn_Reset[43] := BenchUut4.Reset;
   TraceIn_ExtendDone[43] := BenchUut4.ExtendDone;
   TraceIn_ClampDone[43] := BenchUut4.ClampDone;
   TraceIn_ReleaseDone[43] := BenchUut4.ReleaseDone;
   TraceIn_RetractDone[43] := BenchUut4.RetractDone;
   BenchUut4();
   TraceOut_Extend[43] := BenchUut4.Extend;
   TraceOut_Clamp[43] := BenchUut4.Clamp;
   TraceOut_Release[43] := BenchUut4.Release;
   TraceOut_Retract[43] := BenchUut4.Retract;
   TraceOut_Busy[43] := BenchUut4.Busy;
   TraceOut_Done[43] := BenchUut4.Done;
   BenchCalls := BenchCalls + 1;
 44:
   BenchUut4.Start := FALSE;
   BenchUut4.Stop := FALSE;
   BenchUut4.Reset := FALSE;
   BenchUut4.ExtendDone := FALSE;
   BenchUut4.ClampDone := FALSE;
   BenchUut4.ReleaseDone := FALSE;
   BenchUut4.RetractDone := FALSE;
   TraceIn_Start[44] := BenchUut4.Start;
   TraceIn_Stop[44] := BenchUut4.Stop;
   TraceIn_Reset[44] := BenchUut4.Reset;
   TraceIn_ExtendDone[44] := BenchUut4.ExtendDone;
   TraceIn_ClampDone[44] := BenchUut4.ClampDone;
   TraceIn_ReleaseDone[44] := BenchUut4.ReleaseDone;
   TraceIn_RetractDone[44] := BenchUut4.RetractDone;
   BenchUut4();
   TraceOut_Extend[44] := BenchUut4.Extend;
   TraceOut_Clamp[44] := BenchUut4.Clamp;
   TraceOut_Release[44] := BenchUut4.Release;
   TraceOut_Retract[44] := BenchUut4.Retract;
   TraceOut_Busy[44] := BenchUut4.Busy;
   TraceOut_Done[44] := BenchUut4.Done;
   BenchCalls := BenchCalls + 1;
 45:
   BenchUut4.Start := FALSE;
   BenchUut4.Stop := FALSE;
   BenchUut4.Reset := FALSE;
   BenchUut4.ExtendDone := FALSE;
   BenchUut4.ClampDone := FALSE;
   BenchUut4.ReleaseDone := FALSE;
   BenchUut4.RetractDone := FALSE;
   TraceIn_Start[45] := BenchUut4.Start;
   TraceIn_Stop[45] := BenchUut4.Stop;
   TraceIn_Reset[45] := BenchUut4.Reset;
   TraceIn_ExtendDone[45] := BenchUut4.ExtendDone;
   TraceIn_ClampDone[45] := BenchUut4.ClampDone;
   TraceIn_ReleaseDone[45] := BenchUut4.ReleaseDone;
   TraceIn_RetractDone[45] := BenchUut4.RetractDone;
   BenchUut4();
   TraceOut_Extend[45] := BenchUut4.Extend;
   TraceOut_Clamp[45] := BenchUut4.Clamp;
   TraceOut_Release[45] := BenchUut4.Release;
   TraceOut_Retract[45] := BenchUut4.Retract;
   TraceOut_Busy[45] := BenchUut4.Busy;
   TraceOut_Done[45] := BenchUut4.Done;
   BenchCalls := BenchCalls + 1;
 46:
   BenchUut4.Start := FALSE;
   BenchUut4.Stop := FALSE;
   BenchUut4.Reset := FALSE;
   BenchUut4.ExtendDone := FALSE;
   BenchUut4.ClampDone := FALSE;
   BenchUut4.ReleaseDone := FALSE;
   BenchUut4.RetractDone := TRUE;
   TraceIn_Start[46] := BenchUut4.Start;
   TraceIn_Stop[46] := BenchUut4.Stop;
   TraceIn_Reset[46] := BenchUut4.Reset;
   TraceIn_ExtendDone[46] := BenchUut4.ExtendDone;
   TraceIn_ClampDone[46] := BenchUut4.ClampDone;
   TraceIn_ReleaseDone[46] := BenchUut4.ReleaseDone;
   TraceIn_RetractDone[46] := BenchUut4.RetractDone;
   BenchUut4();
   TraceOut_Extend[46] := BenchUut4.Extend;
   TraceOut_Clamp[46] := BenchUut4.Clamp;
   TraceOut_Release[46] := BenchUut4.Release;
   TraceOut_Retract[46] := BenchUut4.Retract;
   TraceOut_Busy[46] := BenchUut4.Busy;
   TraceOut_Done[46] := BenchUut4.Done;
   BenchCalls := BenchCalls + 1;
 47:
   BenchUut4.Start := FALSE;
   BenchUut4.Stop := FALSE;
   BenchUut4.Reset := FALSE;
   BenchUut4.ExtendDone := FALSE;
   BenchUut4.ClampDone := FALSE;
   BenchUut4.ReleaseDone := FALSE;
   BenchUut4.RetractDone := FALSE;
   TraceIn_Start[47] := BenchUut4.Start;
   TraceIn_Stop[47] := BenchUut4.Stop;
   TraceIn_Reset[47] := BenchUut4.Reset;
   TraceIn_ExtendDone[47] := BenchUut4.ExtendDone;
   TraceIn_ClampDone[47] := BenchUut4.ClampDone;
   TraceIn_ReleaseDone[47] := BenchUut4.ReleaseDone;
   TraceIn_RetractDone[47] := BenchUut4.RetractDone;
   BenchUut4();
   TraceOut_Extend[47] := BenchUut4.Extend;
   TraceOut_Clamp[47] := BenchUut4.Clamp;
   TraceOut_Release[47] := BenchUut4.Release;
   TraceOut_Retract[47] := BenchUut4.Retract;
   TraceOut_Busy[47] := BenchUut4.Busy;
   TraceOut_Done[47] := BenchUut4.Done;
   BenchCalls := BenchCalls + 1;
 48:
   BenchUut4.Start := FALSE;
   BenchUut4.Stop := FALSE;
   BenchUut4.Reset := FALSE;
   BenchUut4.ExtendDone := FALSE;
   BenchUut4.ClampDone := FALSE;
   BenchUut4.ReleaseDone := FALSE;
   BenchUut4.RetractDone := FALSE;
   TraceIn_Start[48] := BenchUut4.Start;
   TraceIn_Stop[48] := BenchUut4.Stop;
   TraceIn_Reset[48] := BenchUut4.Reset;
   TraceIn_ExtendDone[48] := BenchUut4.ExtendDone;
   TraceIn_ClampDone[48] := BenchUut4.ClampDone;
   TraceIn_ReleaseDone[48] := BenchUut4.ReleaseDone;
   TraceIn_RetractDone[48] := BenchUut4.RetractDone;
   BenchUut4();
   TraceOut_Extend[48] := BenchUut4.Extend;
   TraceOut_Clamp[48] := BenchUut4.Clamp;
   TraceOut_Release[48] := BenchUut4.Release;
   TraceOut_Retract[48] := BenchUut4.Retract;
   TraceOut_Busy[48] := BenchUut4.Busy;
   TraceOut_Done[48] := BenchUut4.Done;
   BenchCalls := BenchCalls + 1;
 49:
   BenchUut4.Start := FALSE;
   BenchUut4.Stop := FALSE;
   BenchUut4.Reset := FALSE;
   BenchUut4.ExtendDone := FALSE;
   BenchUut4.ClampDone := FALSE;
   BenchUut4.ReleaseDone := FALSE;
   BenchUut4.RetractDone := FALSE;
   TraceIn_Start[49] := BenchUut4.Start;
   TraceIn_Stop[49] := BenchUut4.Stop;
   TraceIn_Reset[49] := BenchUut4.Reset;
   TraceIn_ExtendDone[49] := BenchUut4.ExtendDone;
   TraceIn_ClampDone[49] := BenchUut4.ClampDone;
   TraceIn_ReleaseDone[49] := BenchUut4.ReleaseDone;
   TraceIn_RetractDone[49] := BenchUut4.RetractDone;
   BenchUut4();
   TraceOut_Extend[49] := BenchUut4.Extend;
   TraceOut_Clamp[49] := BenchUut4.Clamp;
   TraceOut_Release[49] := BenchUut4.Release;
   TraceOut_Retract[49] := BenchUut4.Retract;
   TraceOut_Busy[49] := BenchUut4.Busy;
   TraceOut_Done[49] := BenchUut4.Done;
   BenchCalls := BenchCalls + 1;
 50:
   BenchUut4.Start := FALSE;
   BenchUut4.Stop := FALSE;
   BenchUut4.Reset := TRUE;
   BenchUut4.ExtendDone := FALSE;
   BenchUut4.ClampDone := FALSE;
   BenchUut4.ReleaseDone := FALSE;
   BenchUut4.RetractDone := TRUE;
   TraceIn_Start[50] := BenchUut4.Start;
   TraceIn_Stop[50] := BenchUut4.Stop;
   TraceIn_Reset[50] := BenchUut4.Reset;
   TraceIn_ExtendDone[50] := BenchUut4.ExtendDone;
   TraceIn_ClampDone[50] := BenchUut4.ClampDone;
   TraceIn_ReleaseDone[50] := BenchUut4.ReleaseDone;
   TraceIn_RetractDone[50] := BenchUut4.RetractDone;
   BenchUut4();
   TraceOut_Extend[50] := BenchUut4.Extend;
   TraceOut_Clamp[50] := BenchUut4.Clamp;
   TraceOut_Release[50] := BenchUut4.Release;
   TraceOut_Retract[50] := BenchUut4.Retract;
   TraceOut_Busy[50] := BenchUut4.Busy;
   TraceOut_Done[50] := BenchUut4.Done;
   BenchCalls := BenchCalls + 1;
 51:
   BenchUut4.Start := FALSE;
   BenchUut4.Stop := FALSE;
   BenchUut4.Reset := FALSE;
   BenchUut4.ExtendDone := FALSE;
   BenchUut4.ClampDone := FALSE;
   BenchUut4.ReleaseDone := FALSE;
   BenchUut4.RetractDone := TRUE;
   TraceIn_Start[51] := BenchUut4.Start;
   TraceIn_Stop[51] := BenchUut4.Stop;
   TraceIn_Reset[51] := BenchUut4.Reset;
   TraceIn_ExtendDone[51] := BenchUut4.ExtendDone;
   TraceIn_ClampDone[51] := BenchUut4.ClampDone;
   TraceIn_ReleaseDone[51] := BenchUut4.ReleaseDone;
   TraceIn_RetractDone[51] := BenchUut4.RetractDone;
   BenchUut4();
   TraceOut_Extend[51] := BenchUut4.Extend;
   TraceOut_Clamp[51] := BenchUut4.Clamp;
   TraceOut_Release[51] := BenchUut4.Release;
   TraceOut_Retract[51] := BenchUut4.Retract;
   TraceOut_Busy[51] := BenchUut4.Busy;
   TraceOut_Done[51] := BenchUut4.Done;
   BenchCalls := BenchCalls + 1;
 52:
   BenchUut4.Start := TRUE;
   BenchUut4.Stop := FALSE;
   BenchUut4.Reset := FALSE;
   BenchUut4.ExtendDone := FALSE;
   BenchUut4.ClampDone := FALSE;
   BenchUut4.ReleaseDone := FALSE;
   BenchUut4.RetractDone := TRUE;
   TraceIn_Start[52] := BenchUut4.Start;
   TraceIn_Stop[52] := BenchUut4.Stop;
   TraceIn_Reset[52] := BenchUut4.Reset;
   TraceIn_ExtendDone[52] := BenchUut4.ExtendDone;
   TraceIn_ClampDone[52] := BenchUut4.ClampDone;
   TraceIn_ReleaseDone[52] := BenchUut4.ReleaseDone;
   TraceIn_RetractDone[52] := BenchUut4.RetractDone;
   BenchUut4();
   TraceOut_Extend[52] := BenchUut4.Extend;
   TraceOut_Clamp[52] := BenchUut4.Clamp;
   TraceOut_Release[52] := BenchUut4.Release;
   TraceOut_Retract[52] := BenchUut4.Retract;
   TraceOut_Busy[52] := BenchUut4.Busy;
   TraceOut_Done[52] := BenchUut4.Done;
   BenchCalls := BenchCalls + 1;
 53:
   BenchUut4.Start := FALSE;
   BenchUut4.Stop := FALSE;
   BenchUut4.Reset := FALSE;
   BenchUut4.ExtendDone := FALSE;
   BenchUut4.ClampDone := FALSE;
   BenchUut4.ReleaseDone := FALSE;
   BenchUut4.RetractDone := FALSE;
   TraceIn_Start[53] := BenchUut4.Start;
   TraceIn_Stop[53] := BenchUut4.Stop;
   TraceIn_Reset[53] := BenchUut4.Reset;
   TraceIn_ExtendDone[53] := BenchUut4.ExtendDone;
   TraceIn_ClampDone[53] := BenchUut4.ClampDone;
   TraceIn_ReleaseDone[53] := BenchUut4.ReleaseDone;
   TraceIn_RetractDone[53] := BenchUut4.RetractDone;
   BenchUut4();
   TraceOut_Extend[53] := BenchUut4.Extend;
   TraceOut_Clamp[53] := BenchUut4.Clamp;
   TraceOut_Release[53] := BenchUut4.Release;
   TraceOut_Retract[53] := BenchUut4.Retract;
   TraceOut_Busy[53] := BenchUut4.Busy;
   TraceOut_Done[53] := BenchUut4.Done;
   BenchCalls := BenchCalls + 1;
 54:
   BenchUut4.Start := FALSE;
   BenchUut4.Stop := FALSE;
   BenchUut4.Reset := FALSE;
   BenchUut4.ExtendDone := FALSE;
   BenchUut4.ClampDone := FALSE;
   BenchUut4.ReleaseDone := FALSE;
   BenchUut4.RetractDone := FALSE;
   TraceIn_Start[54] := BenchUut4.Start;
   TraceIn_Stop[54] := BenchUut4.Stop;
   TraceIn_Reset[54] := BenchUut4.Reset;
   TraceIn_ExtendDone[54] := BenchUut4.ExtendDone;
   TraceIn_ClampDone[54] := BenchUut4.ClampDone;
   TraceIn_ReleaseDone[54] := BenchUut4.ReleaseDone;
   TraceIn_RetractDone[54] := BenchUut4.RetractDone;
   BenchUut4();
   TraceOut_Extend[54] := BenchUut4.Extend;
   TraceOut_Clamp[54] := BenchUut4.Clamp;
   TraceOut_Release[54] := BenchUut4.Release;
   TraceOut_Retract[54] := BenchUut4.Retract;
   TraceOut_Busy[54] := BenchUut4.Busy;
   TraceOut_Done[54] := BenchUut4.Done;
   BenchCalls := BenchCalls + 1;
 55:
   BenchUut4.Start := FALSE;
   BenchUut4.Stop := FALSE;
   BenchUut4.Reset := FALSE;
   BenchUut4.ExtendDone := TRUE;
   BenchUut4.ClampDone := FALSE;
   BenchUut4.ReleaseDone := FALSE;
   BenchUut4.RetractDone := FALSE;
   TraceIn_Start[55] := BenchUut4.Start;
   TraceIn_Stop[55] := BenchUut4.Stop;
   TraceIn_Reset[55] := BenchUut4.Reset;
   TraceIn_ExtendDone[55] := BenchUut4.ExtendDone;
   TraceIn_ClampDone[55] := BenchUut4.ClampDone;
   TraceIn_ReleaseDone[55] := BenchUut4.ReleaseDone;
   TraceIn_RetractDone[55] := BenchUut4.RetractDone;
   BenchUut4();
   TraceOut_Extend[55] := BenchUut4.Extend;
   TraceOut_Clamp[55] := BenchUut4.Clamp;
   TraceOut_Release[55] := BenchUut4.Release;
   TraceOut_Retract[55] := BenchUut4.Retract;
   TraceOut_Busy[55] := BenchUut4.Busy;
   TraceOut_Done[55] := BenchUut4.Done;
   BenchCalls := BenchCalls + 1;
 56:
   BenchUut4.Start := FALSE;
   BenchUut4.Stop := FALSE;
   BenchUut4.Reset := FALSE;
   BenchUut4.ExtendDone := FALSE;
   BenchUut4.ClampDone := FALSE;
   BenchUut4.ReleaseDone := FALSE;
   BenchUut4.RetractDone := FALSE;
   TraceIn_Start[56] := BenchUut4.Start;
   TraceIn_Stop[56] := BenchUut4.Stop;
   TraceIn_Reset[56] := BenchUut4.Reset;
   TraceIn_ExtendDone[56] := BenchUut4.ExtendDone;
   TraceIn_ClampDone[56] := BenchUut4.ClampDone;
   TraceIn_ReleaseDone[56] := BenchUut4.ReleaseDone;
   TraceIn_RetractDone[56] := BenchUut4.RetractDone;
   BenchUut4();
   TraceOut_Extend[56] := BenchUut4.Extend;
   TraceOut_Clamp[56] := BenchUut4.Clamp;
   TraceOut_Release[56] := BenchUut4.Release;
   TraceOut_Retract[56] := BenchUut4.Retract;
   TraceOut_Busy[56] := BenchUut4.Busy;
   TraceOut_Done[56] := BenchUut4.Done;
   BenchCalls := BenchCalls + 1;
 57:
   BenchUut4.Start := FALSE;
   BenchUut4.Stop := FALSE;
   BenchUut4.Reset := FALSE;
   BenchUut4.ExtendDone := FALSE;
   BenchUut4.ClampDone := FALSE;
   BenchUut4.ReleaseDone := FALSE;
   BenchUut4.RetractDone := FALSE;
   TraceIn_Start[57] := BenchUut4.Start;
   TraceIn_Stop[57] := BenchUut4.Stop;
   TraceIn_Reset[57] := BenchUut4.Reset;
   TraceIn_ExtendDone[57] := BenchUut4.ExtendDone;
   TraceIn_ClampDone[57] := BenchUut4.ClampDone;
   TraceIn_ReleaseDone[57] := BenchUut4.ReleaseDone;
   TraceIn_RetractDone[57] := BenchUut4.RetractDone;
   BenchUut4();
   TraceOut_Extend[57] := BenchUut4.Extend;
   TraceOut_Clamp[57] := BenchUut4.Clamp;
   TraceOut_Release[57] := BenchUut4.Release;
   TraceOut_Retract[57] := BenchUut4.Retract;
   TraceOut_Busy[57] := BenchUut4.Busy;
   TraceOut_Done[57] := BenchUut4.Done;
   BenchCalls := BenchCalls + 1;
 58:
   BenchUut4.Start := FALSE;
   BenchUut4.Stop := FALSE;
   BenchUut4.Reset := FALSE;
   BenchUut4.ExtendDone := FALSE;
   BenchUut4.ClampDone := FALSE;
   BenchUut4.ReleaseDone := FALSE;
   BenchUut4.RetractDone := FALSE;
   TraceIn_Start[58] := BenchUut4.Start;
   TraceIn_Stop[58] := BenchUut4.Stop;
   TraceIn_Reset[58] := BenchUut4.Reset;
   TraceIn_ExtendDone[58] := BenchUut4.ExtendDone;
   TraceIn_ClampDone[58] := BenchUut4.ClampDone;
   TraceIn_ReleaseDone[58] := BenchUut4.ReleaseDone;
   TraceIn_RetractDone[58] := BenchUut4.RetractDone;
   BenchUut4();
   TraceOut_Extend[58] := BenchUut4.Extend;
   TraceOut_Clamp[58] := BenchUut4.Clamp;
   TraceOut_Release[58] := BenchUut4.Release;
   TraceOut_Retract[58] := BenchUut4.Retract;
   TraceOut_Busy[58] := BenchUut4.Busy;
   TraceOut_Done[58] := BenchUut4.Done;
   BenchCalls := BenchCalls + 1;
 59:
   BenchUut4.Start := FALSE;
   BenchUut4.Stop := FALSE;
   BenchUut4.Reset := FALSE;
   BenchUut4.ExtendDone := FALSE;
   BenchUut4.ClampDone := TRUE;
   BenchUut4.ReleaseDone := FALSE;
   BenchUut4.RetractDone := FALSE;
   TraceIn_Start[59] := BenchUut4.Start;
   TraceIn_Stop[59] := BenchUut4.Stop;
   TraceIn_Reset[59] := BenchUut4.Reset;
   TraceIn_ExtendDone[59] := BenchUut4.ExtendDone;
   TraceIn_ClampDone[59] := BenchUut4.ClampDone;
   TraceIn_ReleaseDone[59] := BenchUut4.ReleaseDone;
   TraceIn_RetractDone[59] := BenchUut4.RetractDone;
   BenchUut4();
   TraceOut_Extend[59] := BenchUut4.Extend;
   TraceOut_Clamp[59] := BenchUut4.Clamp;
   TraceOut_Release[59] := BenchUut4.Release;
   TraceOut_Retract[59] := BenchUut4.Retract;
   TraceOut_Busy[59] := BenchUut4.Busy;
   TraceOut_Done[59] := BenchUut4.Done;
   BenchCalls := BenchCalls + 1;
 60:
   BenchUut4.Start := FALSE;
   BenchUut4.Stop := FALSE;
   BenchUut4.Reset := FALSE;
   BenchUut4.ExtendDone := FALSE;
   BenchUut4.ClampDone := FALSE;
   BenchUut4.ReleaseDone := FALSE;
   BenchUut4.RetractDone := FALSE;
   TraceIn_Start[60] := BenchUut4.Start;
   TraceIn_Stop[60] := BenchUut4.Stop;
   TraceIn_Reset[60] := BenchUut4.Reset;
   TraceIn_ExtendDone[60] := BenchUut4.ExtendDone;
   TraceIn_ClampDone[60] := BenchUut4.ClampDone;
   TraceIn_ReleaseDone[60] := BenchUut4.ReleaseDone;
   TraceIn_RetractDone[60] := BenchUut4.RetractDone;
   BenchUut4();
   TraceOut_Extend[60] := BenchUut4.Extend;
   TraceOut_Clamp[60] := BenchUut4.Clamp;
   TraceOut_Release[60] := BenchUut4.Release;
   TraceOut_Retract[60] := BenchUut4.Retract;
   TraceOut_Busy[60] := BenchUut4.Busy;
   TraceOut_Done[60] := BenchUut4.Done;
   BenchCalls := BenchCalls + 1;
 61:
   BenchUut4.Start := FALSE;
   BenchUut4.Stop := FALSE;
   BenchUut4.Reset := FALSE;
   BenchUut4.ExtendDone := FALSE;
   BenchUut4.ClampDone := FALSE;
   BenchUut4.ReleaseDone := FALSE;
   BenchUut4.RetractDone := FALSE;
   TraceIn_Start[61] := BenchUut4.Start;
   TraceIn_Stop[61] := BenchUut4.Stop;
   TraceIn_Reset[61] := BenchUut4.Reset;
   TraceIn_ExtendDone[61] := BenchUut4.ExtendDone;
   TraceIn_ClampDone[61] := BenchUut4.ClampDone;
   TraceIn_ReleaseDone[61] := BenchUut4.ReleaseDone;
   TraceIn_RetractDone[61] := BenchUut4.RetractDone;
   BenchUut4();
   TraceOut_Extend[61] := BenchUut4.Extend;
   TraceOut_Clamp[61] := BenchUut4.Clamp;
   TraceOut_Release[61] := BenchUut4.Release;
   TraceOut_Retract[61] := BenchUut4.Retract;
   TraceOut_Busy[61] := BenchUut4.Busy;
   TraceOut_Done[61] := BenchUut4.Done;
   BenchCalls := BenchCalls + 1;
 62:
   BenchUut4.Start := FALSE;
   BenchUut4.Stop := FALSE;
   BenchUut4.Reset := FALSE;
   BenchUut4.ExtendDone := FALSE;
   BenchUut4.ClampDone := FALSE;
   BenchUut4.ReleaseDone := FALSE;
   BenchUut4.RetractDone := FALSE;
   TraceIn_Start[62] := BenchUut4.Start;
   TraceIn_Stop[62] := BenchUut4.Stop;
   TraceIn_Reset[62] := BenchUut4.Reset;
   TraceIn_ExtendDone[62] := BenchUut4.ExtendDone;
   TraceIn_ClampDone[62] := BenchUut4.ClampDone;
   TraceIn_ReleaseDone[62] := BenchUut4.ReleaseDone;
   TraceIn_RetractDone[62] := BenchUut4.RetractDone;
   BenchUut4();
   TraceOut_Extend[62] := BenchUut4.Extend;
   TraceOut_Clamp[62] := BenchUut4.Clamp;
   TraceOut_Release[62] := BenchUut4.Release;
   TraceOut_Retract[62] := BenchUut4.Retract;
   TraceOut_Busy[62] := BenchUut4.Busy;
   TraceOut_Done[62] := BenchUut4.Done;
   BenchCalls := BenchCalls + 1;
 63:
   BenchUut4.Start := FALSE;
   BenchUut4.Stop := FALSE;
   BenchUut4.Reset := FALSE;
   BenchUut4.ExtendDone := FALSE;
   BenchUut4.ClampDone := FALSE;
   BenchUut4.ReleaseDone := TRUE;
   BenchUut4.RetractDone := FALSE;
   TraceIn_Start[63] := BenchUut4.Start;
   TraceIn_Stop[63] := BenchUut4.Stop;
   TraceIn_Reset[63] := BenchUut4.Reset;
   TraceIn_ExtendDone[63] := BenchUut4.ExtendDone;
   TraceIn_ClampDone[63] := BenchUut4.ClampDone;
   TraceIn_ReleaseDone[63] := BenchUut4.ReleaseDone;
   TraceIn_RetractDone[63] := BenchUut4.RetractDone;
   BenchUut4();
   TraceOut_Extend[63] := BenchUut4.Extend;
   TraceOut_Clamp[63] := BenchUut4.Clamp;
   TraceOut_Release[63] := BenchUut4.Release;
   TraceOut_Retract[63] := BenchUut4.Retract;
   TraceOut_Busy[63] := BenchUut4.Busy;
   TraceOut_Done[63] := BenchUut4.Done;
   BenchCalls := BenchCalls + 1;
 64:
   BenchUut4.Start := FALSE;
   BenchUut4.Stop := FALSE;
   BenchUut4.Reset := FALSE;
   BenchUut4.ExtendDone := FALSE;
   BenchUut4.ClampDone := FALSE;
   BenchUut4.ReleaseDone := FALSE;
   BenchUut4.RetractDone := FALSE;
   TraceIn_Start[64] := BenchUut4.Start;
   TraceIn_Stop[64] := BenchUut4.Stop;
   TraceIn_Reset[64] := BenchUut4.Reset;
   TraceIn_ExtendDone[64] := BenchUut4.ExtendDone;
   TraceIn_ClampDone[64] := BenchUut4.ClampDone;
   TraceIn_ReleaseDone[64] := BenchUut4.ReleaseDone;
   TraceIn_RetractDone[64] := BenchUut4.RetractDone;
   BenchUut4();
   TraceOut_Extend[64] := BenchUut4.Extend;
   TraceOut_Clamp[64] := BenchUut4.Clamp;
   TraceOut_Release[64] := BenchUut4.Release;
   TraceOut_Retract[64] := BenchUut4.Retract;
   TraceOut_Busy[64] := BenchUut4.Busy;
   TraceOut_Done[64] := BenchUut4.Done;
   BenchCalls := BenchCalls + 1;
 65:
   BenchUut4.Start := FALSE;
   BenchUut4.Stop := FALSE;
   BenchUut4.Reset := FALSE;
   BenchUut4.ExtendDone := FALSE;
   BenchUut4.ClampDone := FALSE;
   BenchUut4.ReleaseDone := FALSE;
   BenchUut4.RetractDone := FALSE;
   TraceIn_Start[65] := BenchUut4.Start;
   TraceIn_Stop[65] := BenchUut4.Stop;
   TraceIn_Reset[65] := BenchUut4.Reset;
   TraceIn_ExtendDone[65] := BenchUut4.ExtendDone;
   TraceIn_ClampDone[65] := BenchUut4.ClampDone;
   TraceIn_ReleaseDone[65] := BenchUut4.ReleaseDone;
   TraceIn_RetractDone[65] := BenchUut4.RetractDone;
   BenchUut4();
   TraceOut_Extend[65] := BenchUut4.Extend;
   TraceOut_Clamp[65] := BenchUut4.Clamp;
   TraceOut_Release[65] := BenchUut4.Release;
   TraceOut_Retract[65] := BenchUut4.Retract;
   TraceOut_Busy[65] := BenchUut4.Busy;
   TraceOut_Done[65] := BenchUut4.Done;
   BenchCalls := BenchCalls + 1;
 66:
   BenchUut4.Start := FALSE;
   BenchUut4.Stop := FALSE;
   BenchUut4.Reset := FALSE;
   BenchUut4.ExtendDone := FALSE;
   BenchUut4.ClampDone := FALSE;
   BenchUut4.ReleaseDone := FALSE;
   BenchUut4.RetractDone := FALSE;
   TraceIn_Start[66] := BenchUut4.Start;
   TraceIn_Stop[66] := BenchUut4.Stop;
   TraceIn_Reset[66] := BenchUut4.Reset;
   TraceIn_ExtendDone[66] := BenchUut4.ExtendDone;
   TraceIn_ClampDone[66] := BenchUut4.ClampDone;
   TraceIn_ReleaseDone[66] := BenchUut4.ReleaseDone;
   TraceIn_RetractDone[66] := BenchUut4.RetractDone;
   BenchUut4();
   TraceOut_Extend[66] := BenchUut4.Extend;
   TraceOut_Clamp[66] := BenchUut4.Clamp;
   TraceOut_Release[66] := BenchUut4.Release;
   TraceOut_Retract[66] := BenchUut4.Retract;
   TraceOut_Busy[66] := BenchUut4.Busy;
   TraceOut_Done[66] := BenchUut4.Done;
   BenchCalls := BenchCalls + 1;
 67:
   BenchUut4.Start := FALSE;
   BenchUut4.Stop := FALSE;
   BenchUut4.Reset := FALSE;
   BenchUut4.ExtendDone := FALSE;
   BenchUut4.ClampDone := FALSE;
   BenchUut4.ReleaseDone := FALSE;
   BenchUut4.RetractDone := TRUE;
   TraceIn_Start[67] := BenchUut4.Start;
   TraceIn_Stop[67] := BenchUut4.Stop;
   TraceIn_Reset[67] := BenchUut4.Reset;
   TraceIn_ExtendDone[67] := BenchUut4.ExtendDone;
   TraceIn_ClampDone[67] := BenchUut4.ClampDone;
   TraceIn_ReleaseDone[67] := BenchUut4.ReleaseDone;
   TraceIn_RetractDone[67] := BenchUut4.RetractDone;
   BenchUut4();
   TraceOut_Extend[67] := BenchUut4.Extend;
   TraceOut_Clamp[67] := BenchUut4.Clamp;
   TraceOut_Release[67] := BenchUut4.Release;
   TraceOut_Retract[67] := BenchUut4.Retract;
   TraceOut_Busy[67] := BenchUut4.Busy;
   TraceOut_Done[67] := BenchUut4.Done;
   BenchCalls := BenchCalls + 1;
 68:
   BenchUut4.Start := FALSE;
   BenchUut4.Stop := FALSE;
   BenchUut4.Reset := FALSE;
   BenchUut4.ExtendDone := FALSE;
   BenchUut4.ClampDone := FALSE;
   BenchUut4.ReleaseDone := FALSE;
   BenchUut4.RetractDone := FALSE;
   TraceIn_Start[68] := BenchUut4.Start;
   TraceIn_Stop[68] := BenchUut4.Stop;
   TraceIn_Reset[68] := BenchUut4.Reset;
   TraceIn_ExtendDone[68] := BenchUut4.ExtendDone;
   TraceIn_ClampDone[68] := BenchUut4.ClampDone;
   TraceIn_ReleaseDone[68] := BenchUut4.ReleaseDone;
   TraceIn_RetractDone[68] := BenchUut4.RetractDone;
   BenchUut4();
   TraceOut_Extend[68] := BenchUut4.Extend;
   TraceOut_Clamp[68] := BenchUut4.Clamp;
   TraceOut_Release[68] := BenchUut4.Release;
   TraceOut_Retract[68] := BenchUut4.Retract;
   TraceOut_Busy[68] := BenchUut4.Busy;
   TraceOut_Done[68] := BenchUut4.Done;
   BenchCalls := BenchCalls + 1;
 69:
   BenchUut4.Start := FALSE;
   BenchUut4.Stop := FALSE;
   BenchUut4.Reset := FALSE;
   BenchUut4.ExtendDone := FALSE;
   BenchUut4.ClampDone := FALSE;
   BenchUut4.ReleaseDone := FALSE;
   BenchUut4.RetractDone := FALSE;
   TraceIn_Start[69] := BenchUut4.Start;
   TraceIn_Stop[69] := BenchUut4.Stop;
   TraceIn_Reset[69] := BenchUut4.Reset;
   TraceIn_ExtendDone[69] := BenchUut4.ExtendDone;
   TraceIn_ClampDone[69] := BenchUut4.ClampDone;
   TraceIn_ReleaseDone[69] := BenchUut4.ReleaseDone;
   TraceIn_RetractDone[69] := BenchUut4.RetractDone;
   BenchUut4();
   TraceOut_Extend[69] := BenchUut4.Extend;
   TraceOut_Clamp[69] := BenchUut4.Clamp;
   TraceOut_Release[69] := BenchUut4.Release;
   TraceOut_Retract[69] := BenchUut4.Retract;
   TraceOut_Busy[69] := BenchUut4.Busy;
   TraceOut_Done[69] := BenchUut4.Done;
   BenchCalls := BenchCalls + 1;
 70:
   BenchUut4.Start := FALSE;
   BenchUut4.Stop := FALSE;
   BenchUut4.Reset := FALSE;
   BenchUut4.ExtendDone := FALSE;
   BenchUut4.ClampDone := FALSE;
   BenchUut4.ReleaseDone := FALSE;
   BenchUut4.RetractDone := FALSE;
   TraceIn_Start[70] := BenchUut4.Start;
   TraceIn_Stop[70] := BenchUut4.Stop;
   TraceIn_Reset[70] := BenchUut4.Reset;
   TraceIn_ExtendDone[70] := BenchUut4.ExtendDone;
   TraceIn_ClampDone[70] := BenchUut4.ClampDone;
   TraceIn_ReleaseDone[70] := BenchUut4.ReleaseDone;
   TraceIn_RetractDone[70] := BenchUut4.RetractDone;
   BenchUut4();
   TraceOut_Extend[70] := BenchUut4.Extend;
   TraceOut_Clamp[70] := BenchUut4.Clamp;
   TraceOut_Release[70] := BenchUut4.Release;
   TraceOut_Retract[70] := BenchUut4.Retract;
   TraceOut_Busy[70] := BenchUut4.Busy;
   TraceOut_Done[70] := BenchUut4.Done;
   BenchCalls := BenchCalls + 1;
 71:
   BenchUut5.Start := TRUE;
   BenchUut5.Stop := FALSE;
   BenchUut5.Reset := FALSE;
   BenchUut5.ExtendDone := FALSE;
   BenchUut5.ClampDone := FALSE;
   BenchUut5.ReleaseDone := FALSE;
   BenchUut5.RetractDone := FALSE;
   TraceIn_Start[71] := BenchUut5.Start;
   TraceIn_Stop[71] := BenchUut5.Stop;
   TraceIn_Reset[71] := BenchUut5.Reset;
   TraceIn_ExtendDone[71] := BenchUut5.ExtendDone;
   TraceIn_ClampDone[71] := BenchUut5.ClampDone;
   TraceIn_ReleaseDone[71] := BenchUut5.ReleaseDone;
   TraceIn_RetractDone[71] := BenchUut5.RetractDone;
   BenchUut5();
   TraceOut_Extend[71] := BenchUut5.Extend;
   TraceOut_Clamp[71] := BenchUut5.Clamp;
   TraceOut_Release[71] := BenchUut5.Release;
   TraceOut_Retract[71] := BenchUut5.Retract;
   TraceOut_Busy[71] := BenchUut5.Busy;
   TraceOut_Done[71] := BenchUut5.Done;
   BenchCalls := BenchCalls + 1;
 72:
   BenchUut5.Start := TRUE;
   BenchUut5.Stop := FALSE;
   BenchUut5.Reset := FALSE;
   BenchUut5.ExtendDone := FALSE;
   BenchUut5.ClampDone := FALSE;
   BenchUut5.ReleaseDone := FALSE;
   BenchUut5.RetractDone := TRUE;
   TraceIn_Start[72] := BenchUut5.Start;
   TraceIn_Stop[72] := BenchUut5.Stop;
   TraceIn_Reset[72] := BenchUut5.Reset;
   TraceIn_ExtendDone[72] := BenchUut5.ExtendDone;
   TraceIn_ClampDone[72] := BenchUut5.ClampDone;
   TraceIn_ReleaseDone[72] := BenchUut5.ReleaseDone;
   TraceIn_RetractDone[72] := BenchUut5.RetractDone;
   BenchUut5();
   TraceOut_Extend[72] := BenchUut5.Extend;
   TraceOut_Clamp[72] := BenchUut5.Clamp;
   TraceOut_Release[72] := BenchUut5.Release;
   TraceOut_Retract[72] := BenchUut5.Retract;
   TraceOut_Busy[72] := BenchUut5.Busy;
   TraceOut_Done[72] := BenchUut5.Done;
   BenchCalls := BenchCalls + 1;
 73:
   BenchUut5.Start := FALSE;
   BenchUut5.Stop := FALSE;
   BenchUut5.Reset := FALSE;
   BenchUut5.ExtendDone := FALSE;
   BenchUut5.ClampDone := FALSE;
   BenchUut5.ReleaseDone := FALSE;
   BenchUut5.RetractDone := FALSE;
   TraceIn_Start[73] := BenchUut5.Start;
   TraceIn_Stop[73] := BenchUut5.Stop;
   TraceIn_Reset[73] := BenchUut5.Reset;
   TraceIn_ExtendDone[73] := BenchUut5.ExtendDone;
   TraceIn_ClampDone[73] := BenchUut5.ClampDone;
   TraceIn_ReleaseDone[73] := BenchUut5.ReleaseDone;
   TraceIn_RetractDone[73] := BenchUut5.RetractDone;
   BenchUut5();
   TraceOut_Extend[73] := BenchUut5.Extend;
   TraceOut_Clamp[73] := BenchUut5.Clamp;
   TraceOut_Release[73] := BenchUut5.Release;
   TraceOut_Retract[73] := BenchUut5.Retract;
   TraceOut_Busy[73] := BenchUut5.Busy;
   TraceOut_Done[73] := BenchUut5.Done;
   BenchCalls := BenchCalls + 1;
 74:
   BenchUut5.Start := FALSE;
   BenchUut5.Stop := FALSE;
   BenchUut5.Reset := FALSE;
   BenchUut5.ExtendDone := TRUE;
   BenchUut5.ClampDone := FALSE;
   BenchUut5.ReleaseDone := FALSE;
   BenchUut5.RetractDone := FALSE;
   TraceIn_Start[74] := BenchUut5.Start;
   TraceIn_Stop[74] := BenchUut5.Stop;
   TraceIn_Reset[74] := BenchUut5.Reset;
   TraceIn_ExtendDone[74] := BenchUut5.ExtendDone;
   TraceIn_ClampDone[74] := BenchUut5.ClampDone;
   TraceIn_ReleaseDone[74] := BenchUut5.ReleaseDone;
   TraceIn_RetractDone[74] := BenchUut5.RetractDone;
   BenchUut5();
   TraceOut_Extend[74] := BenchUut5.Extend;
   TraceOut_Clamp[74] := BenchUut5.Clamp;
   TraceOut_Release[74] := BenchUut5.Release;
   TraceOut_Retract[74] := BenchUut5.Retract;
   TraceOut_Busy[74] := BenchUut5.Busy;
   TraceOut_Done[74] := BenchUut5.Done;
   BenchCalls := BenchCalls + 1;
 75:
   BenchUut5.Start := FALSE;
   BenchUut5.Stop := FALSE;
   BenchUut5.Reset := FALSE;
   BenchUut5.ExtendDone := FALSE;
   BenchUut5.ClampDone := TRUE;
   BenchUut5.ReleaseDone := FALSE;
   BenchUut5.RetractDone := FALSE;
   TraceIn_Start[75] := BenchUut5.Start;
   TraceIn_Stop[75] := BenchUut5.Stop;
   TraceIn_Reset[75] := BenchUut5.Reset;
   TraceIn_ExtendDone[75] := BenchUut5.ExtendDone;
   TraceIn_ClampDone[75] := BenchUut5.ClampDone;
   TraceIn_ReleaseDone[75] := BenchUut5.ReleaseDone;
   TraceIn_RetractDone[75] := BenchUut5.RetractDone;
   BenchUut5();
   TraceOut_Extend[75] := BenchUut5.Extend;
   TraceOut_Clamp[75] := BenchUut5.Clamp;
   TraceOut_Release[75] := BenchUut5.Release;
   TraceOut_Retract[75] := BenchUut5.Retract;
   TraceOut_Busy[75] := BenchUut5.Busy;
   TraceOut_Done[75] := BenchUut5.Done;
   BenchCalls := BenchCalls + 1;
 76:
   BenchUut5.Start := FALSE;
   BenchUut5.Stop := FALSE;
   BenchUut5.Reset := FALSE;
   BenchUut5.ExtendDone := FALSE;
   BenchUut5.ClampDone := FALSE;
   BenchUut5.ReleaseDone := TRUE;
   BenchUut5.RetractDone := FALSE;
   TraceIn_Start[76] := BenchUut5.Start;
   TraceIn_Stop[76] := BenchUut5.Stop;
   TraceIn_Reset[76] := BenchUut5.Reset;
   TraceIn_ExtendDone[76] := BenchUut5.ExtendDone;
   TraceIn_ClampDone[76] := BenchUut5.ClampDone;
   TraceIn_ReleaseDone[76] := BenchUut5.ReleaseDone;
   TraceIn_RetractDone[76] := BenchUut5.RetractDone;
   BenchUut5();
   TraceOut_Extend[76] := BenchUut5.Extend;
   TraceOut_Clamp[76] := BenchUut5.Clamp;
   TraceOut_Release[76] := BenchUut5.Release;
   TraceOut_Retract[76] := BenchUut5.Retract;
   TraceOut_Busy[76] := BenchUut5.Busy;
   TraceOut_Done[76] := BenchUut5.Done;
   BenchCalls := BenchCalls + 1;
 77:
   BenchUut5.Start := FALSE;
   BenchUut5.Stop := FALSE;
   BenchUut5.Reset := FALSE;
   BenchUut5.ExtendDone := FALSE;
   BenchUut5.ClampDone := FALSE;
   BenchUut5.ReleaseDone := FALSE;
   BenchUut5.RetractDone := TRUE;
   TraceIn_Start[77] := BenchUut5.Start;
   TraceIn_Stop[77] := BenchUut5.Stop;
   TraceIn_Reset[77] := BenchUut5.Reset;
   TraceIn_ExtendDone[77] := BenchUut5.ExtendDone;
   TraceIn_ClampDone[77] := BenchUut5.ClampDone;
   TraceIn_ReleaseDone[77] := BenchUut5.ReleaseDone;
   TraceIn_RetractDone[77] := BenchUut5.RetractDone;
   BenchUut5();
   TraceOut_Extend[77] := BenchUut5.Extend;
   TraceOut_Clamp[77] := BenchUut5.Clamp;
   TraceOut_Release[77] := BenchUut5.Release;
   TraceOut_Retract[77] := BenchUut5.Retract;
   TraceOut_Busy[77] := BenchUut5.Busy;
   TraceOut_Done[77] := BenchUut5.Done;
   BenchCalls := BenchCalls + 1;
 78:
   BenchUut5.Start := TRUE;
   BenchUut5.Stop := FALSE;
   BenchUut5.Reset := FALSE;
   BenchUut5.ExtendDone := FALSE;
   BenchUut5.ClampDone := FALSE;
   BenchUut5.ReleaseDone := FALSE;
   BenchUut5.RetractDone := FALSE;
   TraceIn_Start[78] := BenchUut5.Start;
   TraceIn_Stop[78] := BenchUut5.Stop;
   TraceIn_Reset[78] := BenchUut5.Reset;
   TraceIn_ExtendDone[78] := BenchUut5.ExtendDone;
   TraceIn_ClampDone[78] := BenchUut5.ClampDone;
   TraceIn_ReleaseDone[78] := BenchUut5.ReleaseDone;
   TraceIn_RetractDone[78] := BenchUut5.RetractDone;
   BenchUut5();
   TraceOut_Extend[78] := BenchUut5.Extend;
   TraceOut_Clamp[78] := BenchUut5.Clamp;
   TraceOut_Release[78] := BenchUut5.Release;
   TraceOut_Retract[78] := BenchUut5.Retract;
   TraceOut_Busy[78] := BenchUut5.Busy;
   TraceOut_Done[78] := BenchUut5.Done;
   BenchCalls := BenchCalls + 1;
 79:
   BenchUut5.Start := FALSE;
   BenchUut5.Stop := FALSE;
   BenchUut5.Reset := TRUE;
   BenchUut5.ExtendDone := FALSE;
   BenchUut5.ClampDone := FALSE;
   BenchUut5.ReleaseDone := FALSE;
   BenchUut5.RetractDone := FALSE;
   TraceIn_Start[79] := BenchUut5.Start;
   TraceIn_Stop[79] := BenchUut5.Stop;
   TraceIn_Reset[79] := BenchUut5.Reset;
   TraceIn_ExtendDone[79] := BenchUut5.ExtendDone;
   TraceIn_ClampDone[79] := BenchUut5.ClampDone;
   TraceIn_ReleaseDone[79] := BenchUut5.ReleaseDone;
   TraceIn_RetractDone[79] := BenchUut5.RetractDone;
   BenchUut5();
   TraceOut_Extend[79] := BenchUut5.Extend;
   TraceOut_Clamp[79] := BenchUut5.Clamp;
   TraceOut_Release[79] := BenchUut5.Release;
   TraceOut_Retract[79] := BenchUut5.Retract;
   TraceOut_Busy[79] := BenchUut5.Busy;
   TraceOut_Done[79] := BenchUut5.Done;
   BenchCalls := BenchCalls + 1;
 80:
   BenchUut5.Start := TRUE;
   BenchUut5.Stop := FALSE;
   BenchUut5.Reset := TRUE;
   BenchUut5.ExtendDone := FALSE;
   BenchUut5.ClampDone := FALSE;
   BenchUut5.ReleaseDone := FALSE;
   BenchUut5.RetractDone := FALSE;
   TraceIn_Start[80] := BenchUut5.Start;
   TraceIn_Stop[80] := BenchUut5.Stop;
   TraceIn_Reset[80] := BenchUut5.Reset;
   TraceIn_ExtendDone[80] := BenchUut5.ExtendDone;
   TraceIn_ClampDone[80] := BenchUut5.ClampDone;
   TraceIn_ReleaseDone[80] := BenchUut5.ReleaseDone;
   TraceIn_RetractDone[80] := BenchUut5.RetractDone;
   BenchUut5();
   TraceOut_Extend[80] := BenchUut5.Extend;
   TraceOut_Clamp[80] := BenchUut5.Clamp;
   TraceOut_Release[80] := BenchUut5.Release;
   TraceOut_Retract[80] := BenchUut5.Retract;
   TraceOut_Busy[80] := BenchUut5.Busy;
   TraceOut_Done[80] := BenchUut5.Done;
   BenchCalls := BenchCalls + 1;
 81:
   BenchUut5.Start := TRUE;
   BenchUut5.Stop := FALSE;
   BenchUut5.Reset := TRUE;
   BenchUut5.ExtendDone := FALSE;
   BenchUut5.ClampDone := FALSE;
   BenchUut5.ReleaseDone := FALSE;
   BenchUut5.RetractDone := FALSE;
   TraceIn_Start[81] := BenchUut5.Start;
   TraceIn_Stop[81] := BenchUut5.Stop;
   TraceIn_Reset[81] := BenchUut5.Reset;
   TraceIn_ExtendDone[81] := BenchUut5.ExtendDone;
   TraceIn_ClampDone[81] := BenchUut5.ClampDone;
   TraceIn_ReleaseDone[81] := BenchUut5.ReleaseDone;
   TraceIn_RetractDone[81] := BenchUut5.RetractDone;
   BenchUut5();
   TraceOut_Extend[81] := BenchUut5.Extend;
   TraceOut_Clamp[81] := BenchUut5.Clamp;
   TraceOut_Release[81] := BenchUut5.Release;
   TraceOut_Retract[81] := BenchUut5.Retract;
   TraceOut_Busy[81] := BenchUut5.Busy;
   TraceOut_Done[81] := BenchUut5.Done;
   BenchCalls := BenchCalls + 1;
 82:
   BenchUut6.Start := TRUE;
   BenchUut6.Stop := FALSE;
   BenchUut6.Reset := FALSE;
   BenchUut6.ExtendDone := FALSE;
   BenchUut6.ClampDone := FALSE;
   BenchUut6.ReleaseDone := FALSE;
   BenchUut6.RetractDone := FALSE;
   TraceIn_Start[82] := BenchUut6.Start;
   TraceIn_Stop[82] := BenchUut6.Stop;
   TraceIn_Reset[82] := BenchUut6.Reset;
   TraceIn_ExtendDone[82] := BenchUut6.ExtendDone;
   TraceIn_ClampDone[82] := BenchUut6.ClampDone;
   TraceIn_ReleaseDone[82] := BenchUut6.ReleaseDone;
   TraceIn_RetractDone[82] := BenchUut6.RetractDone;
   BenchUut6();
   TraceOut_Extend[82] := BenchUut6.Extend;
   TraceOut_Clamp[82] := BenchUut6.Clamp;
   TraceOut_Release[82] := BenchUut6.Release;
   TraceOut_Retract[82] := BenchUut6.Retract;
   TraceOut_Busy[82] := BenchUut6.Busy;
   TraceOut_Done[82] := BenchUut6.Done;
   BenchCalls := BenchCalls + 1;
 83:
   BenchUut6.Start := TRUE;
   BenchUut6.Stop := FALSE;
   BenchUut6.Reset := FALSE;
   BenchUut6.ExtendDone := FALSE;
   BenchUut6.ClampDone := FALSE;
   BenchUut6.ReleaseDone := FALSE;
   BenchUut6.RetractDone := TRUE;
   TraceIn_Start[83] := BenchUut6.Start;
   TraceIn_Stop[83] := BenchUut6.Stop;
   TraceIn_Reset[83] := BenchUut6.Reset;
   TraceIn_ExtendDone[83] := BenchUut6.ExtendDone;
   TraceIn_ClampDone[83] := BenchUut6.ClampDone;
   TraceIn_ReleaseDone[83] := BenchUut6.ReleaseDone;
   TraceIn_RetractDone[83] := BenchUut6.RetractDone;
   BenchUut6();
   TraceOut_Extend[83] := BenchUut6.Extend;
   TraceOut_Clamp[83] := BenchUut6.Clamp;
   TraceOut_Release[83] := BenchUut6.Release;
   TraceOut_Retract[83] := BenchUut6.Retract;
   TraceOut_Busy[83] := BenchUut6.Busy;
   TraceOut_Done[83] := BenchUut6.Done;
   BenchCalls := BenchCalls + 1;
 84:
   BenchUut6.Start := FALSE;
   BenchUut6.Stop := FALSE;
   BenchUut6.Reset := FALSE;
   BenchUut6.ExtendDone := FALSE;
   BenchUut6.ClampDone := FALSE;
   BenchUut6.ReleaseDone := FALSE;
   BenchUut6.RetractDone := FALSE;
   TraceIn_Start[84] := BenchUut6.Start;
   TraceIn_Stop[84] := BenchUut6.Stop;
   TraceIn_Reset[84] := BenchUut6.Reset;
   TraceIn_ExtendDone[84] := BenchUut6.ExtendDone;
   TraceIn_ClampDone[84] := BenchUut6.ClampDone;
   TraceIn_ReleaseDone[84] := BenchUut6.ReleaseDone;
   TraceIn_RetractDone[84] := BenchUut6.RetractDone;
   BenchUut6();
   TraceOut_Extend[84] := BenchUut6.Extend;
   TraceOut_Clamp[84] := BenchUut6.Clamp;
   TraceOut_Release[84] := BenchUut6.Release;
   TraceOut_Retract[84] := BenchUut6.Retract;
   TraceOut_Busy[84] := BenchUut6.Busy;
   TraceOut_Done[84] := BenchUut6.Done;
   BenchCalls := BenchCalls + 1;
 85:
   BenchUut6.Start := FALSE;
   BenchUut6.Stop := FALSE;
   BenchUut6.Reset := FALSE;
   BenchUut6.ExtendDone := TRUE;
   BenchUut6.ClampDone := FALSE;
   BenchUut6.ReleaseDone := FALSE;
   BenchUut6.RetractDone := FALSE;
   TraceIn_Start[85] := BenchUut6.Start;
   TraceIn_Stop[85] := BenchUut6.Stop;
   TraceIn_Reset[85] := BenchUut6.Reset;
   TraceIn_ExtendDone[85] := BenchUut6.ExtendDone;
   TraceIn_ClampDone[85] := BenchUut6.ClampDone;
   TraceIn_ReleaseDone[85] := BenchUut6.ReleaseDone;
   TraceIn_RetractDone[85] := BenchUut6.RetractDone;
   BenchUut6();
   TraceOut_Extend[85] := BenchUut6.Extend;
   TraceOut_Clamp[85] := BenchUut6.Clamp;
   TraceOut_Release[85] := BenchUut6.Release;
   TraceOut_Retract[85] := BenchUut6.Retract;
   TraceOut_Busy[85] := BenchUut6.Busy;
   TraceOut_Done[85] := BenchUut6.Done;
   BenchCalls := BenchCalls + 1;
 86:
   BenchUut6.Start := FALSE;
   BenchUut6.Stop := FALSE;
   BenchUut6.Reset := FALSE;
   BenchUut6.ExtendDone := FALSE;
   BenchUut6.ClampDone := TRUE;
   BenchUut6.ReleaseDone := FALSE;
   BenchUut6.RetractDone := FALSE;
   TraceIn_Start[86] := BenchUut6.Start;
   TraceIn_Stop[86] := BenchUut6.Stop;
   TraceIn_Reset[86] := BenchUut6.Reset;
   TraceIn_ExtendDone[86] := BenchUut6.ExtendDone;
   TraceIn_ClampDone[86] := BenchUut6.ClampDone;
   TraceIn_ReleaseDone[86] := BenchUut6.ReleaseDone;
   TraceIn_RetractDone[86] := BenchUut6.RetractDone;
   BenchUut6();
   TraceOut_Extend[86] := BenchUut6.Extend;
   TraceOut_Clamp[86] := BenchUut6.Clamp;
   TraceOut_Release[86] := BenchUut6.Release;
   TraceOut_Retract[86] := BenchUut6.Retract;
   TraceOut_Busy[86] := BenchUut6.Busy;
   TraceOut_Done[86] := BenchUut6.Done;
   BenchCalls := BenchCalls + 1;
 87:
   BenchUut6.Start := FALSE;
   BenchUut6.Stop := FALSE;
   BenchUut6.Reset := FALSE;
   BenchUut6.ExtendDone := FALSE;
   BenchUut6.ClampDone := FALSE;
   BenchUut6.ReleaseDone := TRUE;
   BenchUut6.RetractDone := FALSE;
   TraceIn_Start[87] := BenchUut6.Start;
   TraceIn_Stop[87] := BenchUut6.Stop;
   TraceIn_Reset[87] := BenchUut6.Reset;
   TraceIn_ExtendDone[87] := BenchUut6.ExtendDone;
   TraceIn_ClampDone[87] := BenchUut6.ClampDone;
   TraceIn_ReleaseDone[87] := BenchUut6.ReleaseDone;
   TraceIn_RetractDone[87] := BenchUut6.RetractDone;
   BenchUut6();
   TraceOut_Extend[87] := BenchUut6.Extend;
   TraceOut_Clamp[87] := BenchUut6.Clamp;
   TraceOut_Release[87] := BenchUut6.Release;
   TraceOut_Retract[87] := BenchUut6.Retract;
   TraceOut_Busy[87] := BenchUut6.Busy;
   TraceOut_Done[87] := BenchUut6.Done;
   BenchCalls := BenchCalls + 1;
 88:
   BenchUut6.Start := FALSE;
   BenchUut6.Stop := FALSE;
   BenchUut6.Reset := FALSE;
   BenchUut6.ExtendDone := FALSE;
   BenchUut6.ClampDone := FALSE;
   BenchUut6.ReleaseDone := FALSE;
   BenchUut6.RetractDone := TRUE;
   TraceIn_Start[88] := BenchUut6.Start;
   TraceIn_Stop[88] := BenchUut6.Stop;
   TraceIn_Reset[88] := BenchUut6.Reset;
   TraceIn_ExtendDone[88] := BenchUut6.ExtendDone;
   TraceIn_ClampDone[88] := BenchUut6.ClampDone;
   TraceIn_ReleaseDone[88] := BenchUut6.ReleaseDone;
   TraceIn_RetractDone[88] := BenchUut6.RetractDone;
   BenchUut6();
   TraceOut_Extend[88] := BenchUut6.Extend;
   TraceOut_Clamp[88] := BenchUut6.Clamp;
   TraceOut_Release[88] := BenchUut6.Release;
   TraceOut_Retract[88] := BenchUut6.Retract;
   TraceOut_Busy[88] := BenchUut6.Busy;
   TraceOut_Done[88] := BenchUut6.Done;
   BenchCalls := BenchCalls + 1;
 89:
   BenchUut6.Start := TRUE;
   BenchUut6.Stop := FALSE;
   BenchUut6.Reset := FALSE;
   BenchUut6.ExtendDone := FALSE;
   BenchUut6.ClampDone := FALSE;
   BenchUut6.ReleaseDone := FALSE;
   BenchUut6.RetractDone := FALSE;
   TraceIn_Start[89] := BenchUut6.Start;
   TraceIn_Stop[89] := BenchUut6.Stop;
   TraceIn_Reset[89] := BenchUut6.Reset;
   TraceIn_ExtendDone[89] := BenchUut6.ExtendDone;
   TraceIn_ClampDone[89] := BenchUut6.ClampDone;
   TraceIn_ReleaseDone[89] := BenchUut6.ReleaseDone;
   TraceIn_RetractDone[89] := BenchUut6.RetractDone;
   BenchUut6();
   TraceOut_Extend[89] := BenchUut6.Extend;
   TraceOut_Clamp[89] := BenchUut6.Clamp;
   TraceOut_Release[89] := BenchUut6.Release;
   TraceOut_Retract[89] := BenchUut6.Retract;
   TraceOut_Busy[89] := BenchUut6.Busy;
   TraceOut_Done[89] := BenchUut6.Done;
   BenchCalls := BenchCalls + 1;
 90:
   BenchUut6.Start := FALSE;
   BenchUut6.Stop := FALSE;
   BenchUut6.Reset := TRUE;
   BenchUut6.ExtendDone := FALSE;
   BenchUut6.ClampDone := FALSE;
   BenchUut6.ReleaseDone := FALSE;
   BenchUut6.RetractDone := FALSE;
   TraceIn_Start[90] := BenchUut6.Start;
   TraceIn_Stop[90] := BenchUut6.Stop;
   TraceIn_Reset[90] := BenchUut6.Reset;
   TraceIn_ExtendDone[90] := BenchUut6.ExtendDone;
   TraceIn_ClampDone[90] := BenchUut6.ClampDone;
   TraceIn_ReleaseDone[90] := BenchUut6.ReleaseDone;
   TraceIn_RetractDone[90] := BenchUut6.RetractDone;
   BenchUut6();
   TraceOut_Extend[90] := BenchUut6.Extend;
   TraceOut_Clamp[90] := BenchUut6.Clamp;
   TraceOut_Release[90] := BenchUut6.Release;
   TraceOut_Retract[90] := BenchUut6.Retract;
   TraceOut_Busy[90] := BenchUut6.Busy;
   TraceOut_Done[90] := BenchUut6.Done;
   BenchCalls := BenchCalls + 1;
 91:
   BenchUut6.Start := FALSE;
   BenchUut6.Stop := TRUE;
   BenchUut6.Reset := TRUE;
   BenchUut6.ExtendDone := FALSE;
   BenchUut6.ClampDone := FALSE;
   BenchUut6.ReleaseDone := FALSE;
   BenchUut6.RetractDone := FALSE;
   TraceIn_Start[91] := BenchUut6.Start;
   TraceIn_Stop[91] := BenchUut6.Stop;
   TraceIn_Reset[91] := BenchUut6.Reset;
   TraceIn_ExtendDone[91] := BenchUut6.ExtendDone;
   TraceIn_ClampDone[91] := BenchUut6.ClampDone;
   TraceIn_ReleaseDone[91] := BenchUut6.ReleaseDone;
   TraceIn_RetractDone[91] := BenchUut6.RetractDone;
   BenchUut6();
   TraceOut_Extend[91] := BenchUut6.Extend;
   TraceOut_Clamp[91] := BenchUut6.Clamp;
   TraceOut_Release[91] := BenchUut6.Release;
   TraceOut_Retract[91] := BenchUut6.Retract;
   TraceOut_Busy[91] := BenchUut6.Busy;
   TraceOut_Done[91] := BenchUut6.Done;
   BenchCalls := BenchCalls + 1;
 92:
   BenchUut6.Start := FALSE;
   BenchUut6.Stop := TRUE;
   BenchUut6.Reset := TRUE;
   BenchUut6.ExtendDone := FALSE;
   BenchUut6.ClampDone := FALSE;
   BenchUut6.ReleaseDone := FALSE;
   BenchUut6.RetractDone := FALSE;
   TraceIn_Start[92] := BenchUut6.Start;
   TraceIn_Stop[92] := BenchUut6.Stop;
   TraceIn_Reset[92] := BenchUut6.Reset;
   TraceIn_ExtendDone[92] := BenchUut6.ExtendDone;
   TraceIn_ClampDone[92] := BenchUut6.ClampDone;
   TraceIn_ReleaseDone[92] := BenchUut6.ReleaseDone;
   TraceIn_RetractDone[92] := BenchUut6.RetractDone;
   BenchUut6();
   TraceOut_Extend[92] := BenchUut6.Extend;
   TraceOut_Clamp[92] := BenchUut6.Clamp;
   TraceOut_Release[92] := BenchUut6.Release;
   TraceOut_Retract[92] := BenchUut6.Retract;
   TraceOut_Busy[92] := BenchUut6.Busy;
   TraceOut_Done[92] := BenchUut6.Done;
   BenchCalls := BenchCalls + 1;
 93:
   BenchUut7.Start := TRUE;
   BenchUut7.Stop := FALSE;
   BenchUut7.Reset := FALSE;
   BenchUut7.ExtendDone := FALSE;
   BenchUut7.ClampDone := FALSE;
   BenchUut7.ReleaseDone := FALSE;
   BenchUut7.RetractDone := FALSE;
   TraceIn_Start[93] := BenchUut7.Start;
   TraceIn_Stop[93] := BenchUut7.Stop;
   TraceIn_Reset[93] := BenchUut7.Reset;
   TraceIn_ExtendDone[93] := BenchUut7.ExtendDone;
   TraceIn_ClampDone[93] := BenchUut7.ClampDone;
   TraceIn_ReleaseDone[93] := BenchUut7.ReleaseDone;
   TraceIn_RetractDone[93] := BenchUut7.RetractDone;
   BenchUut7();
   TraceOut_Extend[93] := BenchUut7.Extend;
   TraceOut_Clamp[93] := BenchUut7.Clamp;
   TraceOut_Release[93] := BenchUut7.Release;
   TraceOut_Retract[93] := BenchUut7.Retract;
   TraceOut_Busy[93] := BenchUut7.Busy;
   TraceOut_Done[93] := BenchUut7.Done;
   BenchCalls := BenchCalls + 1;
 94:
   BenchUut7.Start := TRUE;
   BenchUut7.Stop := FALSE;
   BenchUut7.Reset := FALSE;
   BenchUut7.ExtendDone := FALSE;
   BenchUut7.ClampDone := FALSE;
   BenchUut7.ReleaseDone := FALSE;
   BenchUut7.RetractDone := TRUE;
   TraceIn_Start[94] := BenchUut7.Start;
   TraceIn_Stop[94] := BenchUut7.Stop;
   TraceIn_Reset[94] := BenchUut7.Reset;
   TraceIn_ExtendDone[94] := BenchUut7.ExtendDone;
   TraceIn_ClampDone[94] := BenchUut7.ClampDone;
   TraceIn_ReleaseDone[94] := BenchUut7.ReleaseDone;
   TraceIn_RetractDone[94] := BenchUut7.RetractDone;
   BenchUut7();
   TraceOut_Extend[94] := BenchUut7.Extend;
   TraceOut_Clamp[94] := BenchUut7.Clamp;
   TraceOut_Release[94] := BenchUut7.Release;
   TraceOut_Retract[94] := BenchUut7.Retract;
   TraceOut_Busy[94] := BenchUut7.Busy;
   TraceOut_Done[94] := BenchUut7.Done;
   BenchCalls := BenchCalls + 1;
 95:
   BenchUut7.Start := FALSE;
   BenchUut7.Stop := FALSE;
   BenchUut7.Reset := FALSE;
   BenchUut7.ExtendDone := FALSE;
   BenchUut7.ClampDone := FALSE;
   BenchUut7.ReleaseDone := FALSE;
   BenchUut7.RetractDone := FALSE;
   TraceIn_Start[95] := BenchUut7.Start;
   TraceIn_Stop[95] := BenchUut7.Stop;
   TraceIn_Reset[95] := BenchUut7.Reset;
   TraceIn_ExtendDone[95] := BenchUut7.ExtendDone;
   TraceIn_ClampDone[95] := BenchUut7.ClampDone;
   TraceIn_ReleaseDone[95] := BenchUut7.ReleaseDone;
   TraceIn_RetractDone[95] := BenchUut7.RetractDone;
   BenchUut7();
   TraceOut_Extend[95] := BenchUut7.Extend;
   TraceOut_Clamp[95] := BenchUut7.Clamp;
   TraceOut_Release[95] := BenchUut7.Release;
   TraceOut_Retract[95] := BenchUut7.Retract;
   TraceOut_Busy[95] := BenchUut7.Busy;
   TraceOut_Done[95] := BenchUut7.Done;
   BenchCalls := BenchCalls + 1;
 96:
   BenchUut7.Start := FALSE;
   BenchUut7.Stop := FALSE;
   BenchUut7.Reset := FALSE;
   BenchUut7.ExtendDone := TRUE;
   BenchUut7.ClampDone := FALSE;
   BenchUut7.ReleaseDone := FALSE;
   BenchUut7.RetractDone := FALSE;
   TraceIn_Start[96] := BenchUut7.Start;
   TraceIn_Stop[96] := BenchUut7.Stop;
   TraceIn_Reset[96] := BenchUut7.Reset;
   TraceIn_ExtendDone[96] := BenchUut7.ExtendDone;
   TraceIn_ClampDone[96] := BenchUut7.ClampDone;
   TraceIn_ReleaseDone[96] := BenchUut7.ReleaseDone;
   TraceIn_RetractDone[96] := BenchUut7.RetractDone;
   BenchUut7();
   TraceOut_Extend[96] := BenchUut7.Extend;
   TraceOut_Clamp[96] := BenchUut7.Clamp;
   TraceOut_Release[96] := BenchUut7.Release;
   TraceOut_Retract[96] := BenchUut7.Retract;
   TraceOut_Busy[96] := BenchUut7.Busy;
   TraceOut_Done[96] := BenchUut7.Done;
   BenchCalls := BenchCalls + 1;
 97:
   BenchUut7.Start := FALSE;
   BenchUut7.Stop := FALSE;
   BenchUut7.Reset := FALSE;
   BenchUut7.ExtendDone := FALSE;
   BenchUut7.ClampDone := TRUE;
   BenchUut7.ReleaseDone := FALSE;
   BenchUut7.RetractDone := FALSE;
   TraceIn_Start[97] := BenchUut7.Start;
   TraceIn_Stop[97] := BenchUut7.Stop;
   TraceIn_Reset[97] := BenchUut7.Reset;
   TraceIn_ExtendDone[97] := BenchUut7.ExtendDone;
   TraceIn_ClampDone[97] := BenchUut7.ClampDone;
   TraceIn_ReleaseDone[97] := BenchUut7.ReleaseDone;
   TraceIn_RetractDone[97] := BenchUut7.RetractDone;
   BenchUut7();
   TraceOut_Extend[97] := BenchUut7.Extend;
   TraceOut_Clamp[97] := BenchUut7.Clamp;
   TraceOut_Release[97] := BenchUut7.Release;
   TraceOut_Retract[97] := BenchUut7.Retract;
   TraceOut_Busy[97] := BenchUut7.Busy;
   TraceOut_Done[97] := BenchUut7.Done;
   BenchCalls := BenchCalls + 1;
 98:
   BenchUut7.Start := FALSE;
   BenchUut7.Stop := FALSE;
   BenchUut7.Reset := FALSE;
   BenchUut7.ExtendDone := FALSE;
   BenchUut7.ClampDone := FALSE;
   BenchUut7.ReleaseDone := TRUE;
   BenchUut7.RetractDone := FALSE;
   TraceIn_Start[98] := BenchUut7.Start;
   TraceIn_Stop[98] := BenchUut7.Stop;
   TraceIn_Reset[98] := BenchUut7.Reset;
   TraceIn_ExtendDone[98] := BenchUut7.ExtendDone;
   TraceIn_ClampDone[98] := BenchUut7.ClampDone;
   TraceIn_ReleaseDone[98] := BenchUut7.ReleaseDone;
   TraceIn_RetractDone[98] := BenchUut7.RetractDone;
   BenchUut7();
   TraceOut_Extend[98] := BenchUut7.Extend;
   TraceOut_Clamp[98] := BenchUut7.Clamp;
   TraceOut_Release[98] := BenchUut7.Release;
   TraceOut_Retract[98] := BenchUut7.Retract;
   TraceOut_Busy[98] := BenchUut7.Busy;
   TraceOut_Done[98] := BenchUut7.Done;
   BenchCalls := BenchCalls + 1;
 99:
   BenchUut7.Start := FALSE;
   BenchUut7.Stop := FALSE;
   BenchUut7.Reset := FALSE;
   BenchUut7.ExtendDone := FALSE;
   BenchUut7.ClampDone := FALSE;
   BenchUut7.ReleaseDone := FALSE;
   BenchUut7.RetractDone := TRUE;
   TraceIn_Start[99] := BenchUut7.Start;
   TraceIn_Stop[99] := BenchUut7.Stop;
   TraceIn_Reset[99] := BenchUut7.Reset;
   TraceIn_ExtendDone[99] := BenchUut7.ExtendDone;
   TraceIn_ClampDone[99] := BenchUut7.ClampDone;
   TraceIn_ReleaseDone[99] := BenchUut7.ReleaseDone;
   TraceIn_RetractDone[99] := BenchUut7.RetractDone;
   BenchUut7();
   TraceOut_Extend[99] := BenchUut7.Extend;
   TraceOut_Clamp[99] := BenchUut7.Clamp;
   TraceOut_Release[99] := BenchUut7.Release;
   TraceOut_Retract[99] := BenchUut7.Retract;
   TraceOut_Busy[99] := BenchUut7.Busy;
   TraceOut_Done[99] := BenchUut7.Done;
   BenchCalls := BenchCalls + 1;
 100:
   BenchUut7.Start := TRUE;
   BenchUut7.Stop := FALSE;
   BenchUut7.Reset := FALSE;
   BenchUut7.ExtendDone := FALSE;
   BenchUut7.ClampDone := FALSE;
   BenchUut7.ReleaseDone := FALSE;
   BenchUut7.RetractDone := FALSE;
   TraceIn_Start[100] := BenchUut7.Start;
   TraceIn_Stop[100] := BenchUut7.Stop;
   TraceIn_Reset[100] := BenchUut7.Reset;
   TraceIn_ExtendDone[100] := BenchUut7.ExtendDone;
   TraceIn_ClampDone[100] := BenchUut7.ClampDone;
   TraceIn_ReleaseDone[100] := BenchUut7.ReleaseDone;
   TraceIn_RetractDone[100] := BenchUut7.RetractDone;
   BenchUut7();
   TraceOut_Extend[100] := BenchUut7.Extend;
   TraceOut_Clamp[100] := BenchUut7.Clamp;
   TraceOut_Release[100] := BenchUut7.Release;
   TraceOut_Retract[100] := BenchUut7.Retract;
   TraceOut_Busy[100] := BenchUut7.Busy;
   TraceOut_Done[100] := BenchUut7.Done;
   BenchCalls := BenchCalls + 1;
 101:
   BenchUut7.Start := FALSE;
   BenchUut7.Stop := FALSE;
   BenchUut7.Reset := TRUE;
   BenchUut7.ExtendDone := FALSE;
   BenchUut7.ClampDone := FALSE;
   BenchUut7.ReleaseDone := FALSE;
   BenchUut7.RetractDone := FALSE;
   TraceIn_Start[101] := BenchUut7.Start;
   TraceIn_Stop[101] := BenchUut7.Stop;
   TraceIn_Reset[101] := BenchUut7.Reset;
   TraceIn_ExtendDone[101] := BenchUut7.ExtendDone;
   TraceIn_ClampDone[101] := BenchUut7.ClampDone;
   TraceIn_ReleaseDone[101] := BenchUut7.ReleaseDone;
   TraceIn_RetractDone[101] := BenchUut7.RetractDone;
   BenchUut7();
   TraceOut_Extend[101] := BenchUut7.Extend;
   TraceOut_Clamp[101] := BenchUut7.Clamp;
   TraceOut_Release[101] := BenchUut7.Release;
   TraceOut_Retract[101] := BenchUut7.Retract;
   TraceOut_Busy[101] := BenchUut7.Busy;
   TraceOut_Done[101] := BenchUut7.Done;
   BenchCalls := BenchCalls + 1;
 102:
   BenchUut7.Start := FALSE;
   BenchUut7.Stop := FALSE;
   BenchUut7.Reset := FALSE;
   BenchUut7.ExtendDone := FALSE;
   BenchUut7.ClampDone := FALSE;
   BenchUut7.ReleaseDone := FALSE;
   BenchUut7.RetractDone := FALSE;
   TraceIn_Start[102] := BenchUut7.Start;
   TraceIn_Stop[102] := BenchUut7.Stop;
   TraceIn_Reset[102] := BenchUut7.Reset;
   TraceIn_ExtendDone[102] := BenchUut7.ExtendDone;
   TraceIn_ClampDone[102] := BenchUut7.ClampDone;
   TraceIn_ReleaseDone[102] := BenchUut7.ReleaseDone;
   TraceIn_RetractDone[102] := BenchUut7.RetractDone;
   BenchUut7();
   TraceOut_Extend[102] := BenchUut7.Extend;
   TraceOut_Clamp[102] := BenchUut7.Clamp;
   TraceOut_Release[102] := BenchUut7.Release;
   TraceOut_Retract[102] := BenchUut7.Retract;
   TraceOut_Busy[102] := BenchUut7.Busy;
   TraceOut_Done[102] := BenchUut7.Done;
   BenchCalls := BenchCalls + 1;
 103:
   BenchUut7.Start := FALSE;
   BenchUut7.Stop := FALSE;
   BenchUut7.Reset := FALSE;
   BenchUut7.ExtendDone := FALSE;
   BenchUut7.ClampDone := FALSE;
   BenchUut7.ReleaseDone := FALSE;
   BenchUut7.RetractDone := FALSE;
   TraceIn_Start[103] := BenchUut7.Start;
   TraceIn_Stop[103] := BenchUut7.Stop;
   TraceIn_Reset[103] := BenchUut7.Reset;
   TraceIn_ExtendDone[103] := BenchUut7.ExtendDone;
   TraceIn_ClampDone[103] := BenchUut7.ClampDone;
   TraceIn_ReleaseDone[103] := BenchUut7.ReleaseDone;
   TraceIn_RetractDone[103] := BenchUut7.RetractDone;
   BenchUut7();
   TraceOut_Extend[103] := BenchUut7.Extend;
   TraceOut_Clamp[103] := BenchUut7.Clamp;
   TraceOut_Release[103] := BenchUut7.Release;
   TraceOut_Retract[103] := BenchUut7.Retract;
   TraceOut_Busy[103] := BenchUut7.Busy;
   TraceOut_Done[103] := BenchUut7.Done;
   BenchCalls := BenchCalls + 1;
 104:
   BenchUut8.Start := TRUE;
   BenchUut8.Stop := FALSE;
   BenchUut8.Reset := FALSE;
   BenchUut8.ExtendDone := FALSE;
   BenchUut8.ClampDone := FALSE;
   BenchUut8.ReleaseDone := FALSE;
   BenchUut8.RetractDone := FALSE;
   TraceIn_Start[104] := BenchUut8.Start;
   TraceIn_Stop[104] := BenchUut8.Stop;
   TraceIn_Reset[104] := BenchUut8.Reset;
   TraceIn_ExtendDone[104] := BenchUut8.ExtendDone;
   TraceIn_ClampDone[104] := BenchUut8.ClampDone;
   TraceIn_ReleaseDone[104] := BenchUut8.ReleaseDone;
   TraceIn_RetractDone[104] := BenchUut8.RetractDone;
   BenchUut8();
   TraceOut_Extend[104] := BenchUut8.Extend;
   TraceOut_Clamp[104] := BenchUut8.Clamp;
   TraceOut_Release[104] := BenchUut8.Release;
   TraceOut_Retract[104] := BenchUut8.Retract;
   TraceOut_Busy[104] := BenchUut8.Busy;
   TraceOut_Done[104] := BenchUut8.Done;
   BenchCalls := BenchCalls + 1;
 105:
   BenchUut8.Start := TRUE;
   BenchUut8.Stop := FALSE;
   BenchUut8.Reset := FALSE;
   BenchUut8.ExtendDone := FALSE;
   BenchUut8.ClampDone := FALSE;
   BenchUut8.ReleaseDone := FALSE;
   BenchUut8.RetractDone := TRUE;
   TraceIn_Start[105] := BenchUut8.Start;
   TraceIn_Stop[105] := BenchUut8.Stop;
   TraceIn_Reset[105] := BenchUut8.Reset;
   TraceIn_ExtendDone[105] := BenchUut8.ExtendDone;
   TraceIn_ClampDone[105] := BenchUut8.ClampDone;
   TraceIn_ReleaseDone[105] := BenchUut8.ReleaseDone;
   TraceIn_RetractDone[105] := BenchUut8.RetractDone;
   BenchUut8();
   TraceOut_Extend[105] := BenchUut8.Extend;
   TraceOut_Clamp[105] := BenchUut8.Clamp;
   TraceOut_Release[105] := BenchUut8.Release;
   TraceOut_Retract[105] := BenchUut8.Retract;
   TraceOut_Busy[105] := BenchUut8.Busy;
   TraceOut_Done[105] := BenchUut8.Done;
   BenchCalls := BenchCalls + 1;
 106:
   BenchUut8.Start := FALSE;
   BenchUut8.Stop := FALSE;
   BenchUut8.Reset := FALSE;
   BenchUut8.ExtendDone := FALSE;
   BenchUut8.ClampDone := FALSE;
   BenchUut8.ReleaseDone := FALSE;
   BenchUut8.RetractDone := FALSE;
   TraceIn_Start[106] := BenchUut8.Start;
   TraceIn_Stop[106] := BenchUut8.Stop;
   TraceIn_Reset[106] := BenchUut8.Reset;
   TraceIn_ExtendDone[106] := BenchUut8.ExtendDone;
   TraceIn_ClampDone[106] := BenchUut8.ClampDone;
   TraceIn_ReleaseDone[106] := BenchUut8.ReleaseDone;
   TraceIn_RetractDone[106] := BenchUut8.RetractDone;
   BenchUut8();
   TraceOut_Extend[106] := BenchUut8.Extend;
   TraceOut_Clamp[106] := BenchUut8.Clamp;
   TraceOut_Release[106] := BenchUut8.Release;
   TraceOut_Retract[106] := BenchUut8.Retract;
   TraceOut_Busy[106] := BenchUut8.Busy;
   TraceOut_Done[106] := BenchUut8.Done;
   BenchCalls := BenchCalls + 1;
 107:
   BenchUut8.Start := FALSE;
   BenchUut8.Stop := FALSE;
   BenchUut8.Reset := FALSE;
   BenchUut8.ExtendDone := TRUE;
   BenchUut8.ClampDone := FALSE;
   BenchUut8.ReleaseDone := FALSE;
   BenchUut8.RetractDone := FALSE;
   TraceIn_Start[107] := BenchUut8.Start;
   TraceIn_Stop[107] := BenchUut8.Stop;
   TraceIn_Reset[107] := BenchUut8.Reset;
   TraceIn_ExtendDone[107] := BenchUut8.ExtendDone;
   TraceIn_ClampDone[107] := BenchUut8.ClampDone;
   TraceIn_ReleaseDone[107] := BenchUut8.ReleaseDone;
   TraceIn_RetractDone[107] := BenchUut8.RetractDone;
   BenchUut8();
   TraceOut_Extend[107] := BenchUut8.Extend;
   TraceOut_Clamp[107] := BenchUut8.Clamp;
   TraceOut_Release[107] := BenchUut8.Release;
   TraceOut_Retract[107] := BenchUut8.Retract;
   TraceOut_Busy[107] := BenchUut8.Busy;
   TraceOut_Done[107] := BenchUut8.Done;
   BenchCalls := BenchCalls + 1;
 108:
   BenchUut8.Start := FALSE;
   BenchUut8.Stop := FALSE;
   BenchUut8.Reset := FALSE;
   BenchUut8.ExtendDone := FALSE;
   BenchUut8.ClampDone := TRUE;
   BenchUut8.ReleaseDone := FALSE;
   BenchUut8.RetractDone := FALSE;
   TraceIn_Start[108] := BenchUut8.Start;
   TraceIn_Stop[108] := BenchUut8.Stop;
   TraceIn_Reset[108] := BenchUut8.Reset;
   TraceIn_ExtendDone[108] := BenchUut8.ExtendDone;
   TraceIn_ClampDone[108] := BenchUut8.ClampDone;
   TraceIn_ReleaseDone[108] := BenchUut8.ReleaseDone;
   TraceIn_RetractDone[108] := BenchUut8.RetractDone;
   BenchUut8();
   TraceOut_Extend[108] := BenchUut8.Extend;
   TraceOut_Clamp[108] := BenchUut8.Clamp;
   TraceOut_Release[108] := BenchUut8.Release;
   TraceOut_Retract[108] := BenchUut8.Retract;
   TraceOut_Busy[108] := BenchUut8.Busy;
   TraceOut_Done[108] := BenchUut8.Done;
   BenchCalls := BenchCalls + 1;
 109:
   BenchUut8.Start := FALSE;
   BenchUut8.Stop := FALSE;
   BenchUut8.Reset := FALSE;
   BenchUut8.ExtendDone := FALSE;
   BenchUut8.ClampDone := FALSE;
   BenchUut8.ReleaseDone := TRUE;
   BenchUut8.RetractDone := FALSE;
   TraceIn_Start[109] := BenchUut8.Start;
   TraceIn_Stop[109] := BenchUut8.Stop;
   TraceIn_Reset[109] := BenchUut8.Reset;
   TraceIn_ExtendDone[109] := BenchUut8.ExtendDone;
   TraceIn_ClampDone[109] := BenchUut8.ClampDone;
   TraceIn_ReleaseDone[109] := BenchUut8.ReleaseDone;
   TraceIn_RetractDone[109] := BenchUut8.RetractDone;
   BenchUut8();
   TraceOut_Extend[109] := BenchUut8.Extend;
   TraceOut_Clamp[109] := BenchUut8.Clamp;
   TraceOut_Release[109] := BenchUut8.Release;
   TraceOut_Retract[109] := BenchUut8.Retract;
   TraceOut_Busy[109] := BenchUut8.Busy;
   TraceOut_Done[109] := BenchUut8.Done;
   BenchCalls := BenchCalls + 1;
 110:
   BenchUut8.Start := FALSE;
   BenchUut8.Stop := FALSE;
   BenchUut8.Reset := FALSE;
   BenchUut8.ExtendDone := FALSE;
   BenchUut8.ClampDone := FALSE;
   BenchUut8.ReleaseDone := FALSE;
   BenchUut8.RetractDone := TRUE;
   TraceIn_Start[110] := BenchUut8.Start;
   TraceIn_Stop[110] := BenchUut8.Stop;
   TraceIn_Reset[110] := BenchUut8.Reset;
   TraceIn_ExtendDone[110] := BenchUut8.ExtendDone;
   TraceIn_ClampDone[110] := BenchUut8.ClampDone;
   TraceIn_ReleaseDone[110] := BenchUut8.ReleaseDone;
   TraceIn_RetractDone[110] := BenchUut8.RetractDone;
   BenchUut8();
   TraceOut_Extend[110] := BenchUut8.Extend;
   TraceOut_Clamp[110] := BenchUut8.Clamp;
   TraceOut_Release[110] := BenchUut8.Release;
   TraceOut_Retract[110] := BenchUut8.Retract;
   TraceOut_Busy[110] := BenchUut8.Busy;
   TraceOut_Done[110] := BenchUut8.Done;
   BenchCalls := BenchCalls + 1;
 111:
   BenchUut8.Start := TRUE;
   BenchUut8.Stop := FALSE;
   BenchUut8.Reset := FALSE;
   BenchUut8.ExtendDone := FALSE;
   BenchUut8.ClampDone := FALSE;
   BenchUut8.ReleaseDone := FALSE;
   BenchUut8.RetractDone := FALSE;
   TraceIn_Start[111] := BenchUut8.Start;
   TraceIn_Stop[111] := BenchUut8.Stop;
   TraceIn_Reset[111] := BenchUut8.Reset;
   TraceIn_ExtendDone[111] := BenchUut8.ExtendDone;
   TraceIn_ClampDone[111] := BenchUut8.ClampDone;
   TraceIn_ReleaseDone[111] := BenchUut8.ReleaseDone;
   TraceIn_RetractDone[111] := BenchUut8.RetractDone;
   BenchUut8();
   TraceOut_Extend[111] := BenchUut8.Extend;
   TraceOut_Clamp[111] := BenchUut8.Clamp;
   TraceOut_Release[111] := BenchUut8.Release;
   TraceOut_Retract[111] := BenchUut8.Retract;
   TraceOut_Busy[111] := BenchUut8.Busy;
   TraceOut_Done[111] := BenchUut8.Done;
   BenchCalls := BenchCalls + 1;
 112:
   BenchUut8.Start := FALSE;
   BenchUut8.Stop := FALSE;
   BenchUut8.Reset := TRUE;
   BenchUut8.ExtendDone := FALSE;
   BenchUut8.ClampDone := FALSE;
   BenchUut8.ReleaseDone := FALSE;
   BenchUut8.RetractDone := FALSE;
   TraceIn_Start[112] := BenchUut8.Start;
   TraceIn_Stop[112] := BenchUut8.Stop;
   TraceIn_Reset[112] := BenchUut8.Reset;
   TraceIn_ExtendDone[112] := BenchUut8.ExtendDone;
   TraceIn_ClampDone[112] := BenchUut8.ClampDone;
   TraceIn_ReleaseDone[112] := BenchUut8.ReleaseDone;
   TraceIn_RetractDone[112] := BenchUut8.RetractDone;
   BenchUut8();
   TraceOut_Extend[112] := BenchUut8.Extend;
   TraceOut_Clamp[112] := BenchUut8.Clamp;
   TraceOut_Release[112] := BenchUut8.Release;
   TraceOut_Retract[112] := BenchUut8.Retract;
   TraceOut_Busy[112] := BenchUut8.Busy;
   TraceOut_Done[112] := BenchUut8.Done;
   BenchCalls := BenchCalls + 1;
 113:
   BenchUut8.Start := FALSE;
   BenchUut8.Stop := FALSE;
   BenchUut8.Reset := TRUE;
   BenchUut8.ExtendDone := TRUE;
   BenchUut8.ClampDone := FALSE;
   BenchUut8.ReleaseDone := FALSE;
   BenchUut8.RetractDone := FALSE;
   TraceIn_Start[113] := BenchUut8.Start;
   TraceIn_Stop[113] := BenchUut8.Stop;
   TraceIn_Reset[113] := BenchUut8.Reset;
   TraceIn_ExtendDone[113] := BenchUut8.ExtendDone;
   TraceIn_ClampDone[113] := BenchUut8.ClampDone;
   TraceIn_ReleaseDone[113] := BenchUut8.ReleaseDone;
   TraceIn_RetractDone[113] := BenchUut8.RetractDone;
   BenchUut8();
   TraceOut_Extend[113] := BenchUut8.Extend;
   TraceOut_Clamp[113] := BenchUut8.Clamp;
   TraceOut_Release[113] := BenchUut8.Release;
   TraceOut_Retract[113] := BenchUut8.Retract;
   TraceOut_Busy[113] := BenchUut8.Busy;
   TraceOut_Done[113] := BenchUut8.Done;
   BenchCalls := BenchCalls + 1;
 114:
   BenchUut8.Start := FALSE;
   BenchUut8.Stop := FALSE;
   BenchUut8.Reset := TRUE;
   BenchUut8.ExtendDone := TRUE;
   BenchUut8.ClampDone := FALSE;
   BenchUut8.ReleaseDone := FALSE;
   BenchUut8.RetractDone := FALSE;
   TraceIn_Start[114] := BenchUut8.Start;
   TraceIn_Stop[114] := BenchUut8.Stop;
   TraceIn_Reset[114] := BenchUut8.Reset;
   TraceIn_ExtendDone[114] := BenchUut8.ExtendDone;
   TraceIn_ClampDone[114] := BenchUut8.ClampDone;
   TraceIn_ReleaseDone[114] := BenchUut8.ReleaseDone;
   TraceIn_RetractDone[114] := BenchUut8.RetractDone;
   BenchUut8();
   TraceOut_Extend[114] := BenchUut8.Extend;
   TraceOut_Clamp[114] := BenchUut8.Clamp;
   TraceOut_Release[114] := BenchUut8.Release;
   TraceOut_Retract[114] := BenchUut8.Retract;
   TraceOut_Busy[114] := BenchUut8.Busy;
   TraceOut_Done[114] := BenchUut8.Done;
   BenchCalls := BenchCalls + 1;
 115:
   BenchUut9.Start := TRUE;
   BenchUut9.Stop := FALSE;
   BenchUut9.Reset := FALSE;
   BenchUut9.ExtendDone := FALSE;
   BenchUut9.ClampDone := FALSE;
   BenchUut9.ReleaseDone := FALSE;
   BenchUut9.RetractDone := FALSE;
   TraceIn_Start[115] := BenchUut9.Start;
   TraceIn_Stop[115] := BenchUut9.Stop;
   TraceIn_Reset[115] := BenchUut9.Reset;
   TraceIn_ExtendDone[115] := BenchUut9.ExtendDone;
   TraceIn_ClampDone[115] := BenchUut9.ClampDone;
   TraceIn_ReleaseDone[115] := BenchUut9.ReleaseDone;
   TraceIn_RetractDone[115] := BenchUut9.RetractDone;
   BenchUut9();
   TraceOut_Extend[115] := BenchUut9.Extend;
   TraceOut_Clamp[115] := BenchUut9.Clamp;
   TraceOut_Release[115] := BenchUut9.Release;
   TraceOut_Retract[115] := BenchUut9.Retract;
   TraceOut_Busy[115] := BenchUut9.Busy;
   TraceOut_Done[115] := BenchUut9.Done;
   BenchCalls := BenchCalls + 1;
 116:
   BenchUut9.Start := TRUE;
   BenchUut9.Stop := FALSE;
   BenchUut9.Reset := FALSE;
   BenchUut9.ExtendDone := FALSE;
   BenchUut9.ClampDone := FALSE;
   BenchUut9.ReleaseDone := FALSE;
   BenchUut9.RetractDone := TRUE;
   TraceIn_Start[116] := BenchUut9.Start;
   TraceIn_Stop[116] := BenchUut9.Stop;
   TraceIn_Reset[116] := BenchUut9.Reset;
   TraceIn_ExtendDone[116] := BenchUut9.ExtendDone;
   TraceIn_ClampDone[116] := BenchUut9.ClampDone;
   TraceIn_ReleaseDone[116] := BenchUut9.ReleaseDone;
   TraceIn_RetractDone[116] := BenchUut9.RetractDone;
   BenchUut9();
   TraceOut_Extend[116] := BenchUut9.Extend;
   TraceOut_Clamp[116] := BenchUut9.Clamp;
   TraceOut_Release[116] := BenchUut9.Release;
   TraceOut_Retract[116] := BenchUut9.Retract;
   TraceOut_Busy[116] := BenchUut9.Busy;
   TraceOut_Done[116] := BenchUut9.Done;
   BenchCalls := BenchCalls + 1;
 117:
   BenchUut9.Start := FALSE;
   BenchUut9.Stop := FALSE;
   BenchUut9.Reset := FALSE;
   BenchUut9.ExtendDone := FALSE;
   BenchUut9.ClampDone := FALSE;
   BenchUut9.ReleaseDone := FALSE;
   BenchUut9.RetractDone := FALSE;
   TraceIn_Start[117] := BenchUut9.Start;
   TraceIn_Stop[117] := BenchUut9.Stop;
   TraceIn_Reset[117] := BenchUut9.Reset;
   TraceIn_ExtendDone[117] := BenchUut9.ExtendDone;
   TraceIn_ClampDone[117] := BenchUut9.ClampDone;
   TraceIn_ReleaseDone[117] := BenchUut9.ReleaseDone;
   TraceIn_RetractDone[117] := BenchUut9.RetractDone;
   BenchUut9();
   TraceOut_Extend[117] := BenchUut9.Extend;
   TraceOut_Clamp[117] := BenchUut9.Clamp;
   TraceOut_Release[117] := BenchUut9.Release;
   TraceOut_Retract[117] := BenchUut9.Retract;
   TraceOut_Busy[117] := BenchUut9.Busy;
   TraceOut_Done[117] := BenchUut9.Done;
   BenchCalls := BenchCalls + 1;
 118:
   BenchUut9.Start := FALSE;
   BenchUut9.Stop := FALSE;
   BenchUut9.Reset := FALSE;
   BenchUut9.ExtendDone := TRUE;
   BenchUut9.ClampDone := FALSE;
   BenchUut9.ReleaseDone := FALSE;
   BenchUut9.RetractDone := FALSE;
   TraceIn_Start[118] := BenchUut9.Start;
   TraceIn_Stop[118] := BenchUut9.Stop;
   TraceIn_Reset[118] := BenchUut9.Reset;
   TraceIn_ExtendDone[118] := BenchUut9.ExtendDone;
   TraceIn_ClampDone[118] := BenchUut9.ClampDone;
   TraceIn_ReleaseDone[118] := BenchUut9.ReleaseDone;
   TraceIn_RetractDone[118] := BenchUut9.RetractDone;
   BenchUut9();
   TraceOut_Extend[118] := BenchUut9.Extend;
   TraceOut_Clamp[118] := BenchUut9.Clamp;
   TraceOut_Release[118] := BenchUut9.Release;
   TraceOut_Retract[118] := BenchUut9.Retract;
   TraceOut_Busy[118] := BenchUut9.Busy;
   TraceOut_Done[118] := BenchUut9.Done;
   BenchCalls := BenchCalls + 1;
 119:
   BenchUut9.Start := FALSE;
   BenchUut9.Stop := FALSE;
   BenchUut9.Reset := FALSE;
   BenchUut9.ExtendDone := FALSE;
   BenchUut9.ClampDone := TRUE;
   BenchUut9.ReleaseDone := FALSE;
   BenchUut9.RetractDone := FALSE;
   TraceIn_Start[119] := BenchUut9.Start;
   TraceIn_Stop[119] := BenchUut9.Stop;
   TraceIn_Reset[119] := BenchUut9.Reset;
   TraceIn_ExtendDone[119] := BenchUut9.ExtendDone;
   TraceIn_ClampDone[119] := BenchUut9.ClampDone;
   TraceIn_ReleaseDone[119] := BenchUut9.ReleaseDone;
   TraceIn_RetractDone[119] := BenchUut9.RetractDone;
   BenchUut9();
   TraceOut_Extend[119] := BenchUut9.Extend;
   TraceOut_Clamp[119] := BenchUut9.Clamp;
   TraceOut_Release[119] := BenchUut9.Release;
   TraceOut_Retract[119] := BenchUut9.Retract;
   TraceOut_Busy[119] := BenchUut9.Busy;
   TraceOut_Done[119] := BenchUut9.Done;
   BenchCalls := BenchCalls + 1;
 120:
   BenchUut9.Start := FALSE;
   BenchUut9.Stop := FALSE;
   BenchUut9.Reset := FALSE;
   BenchUut9.ExtendDone := FALSE;
   BenchUut9.ClampDone := FALSE;
   BenchUut9.ReleaseDone := TRUE;
   BenchUut9.RetractDone := FALSE;
   TraceIn_Start[120] := BenchUut9.Start;
   TraceIn_Stop[120] := BenchUut9.Stop;
   TraceIn_Reset[120] := BenchUut9.Reset;
   TraceIn_ExtendDone[120] := BenchUut9.ExtendDone;
   TraceIn_ClampDone[120] := BenchUut9.ClampDone;
   TraceIn_ReleaseDone[120] := BenchUut9.ReleaseDone;
   TraceIn_RetractDone[120] := BenchUut9.RetractDone;
   BenchUut9();
   TraceOut_Extend[120] := BenchUut9.Extend;
   TraceOut_Clamp[120] := BenchUut9.Clamp;
   TraceOut_Release[120] := BenchUut9.Release;
   TraceOut_Retract[120] := BenchUut9.Retract;
   TraceOut_Busy[120] := BenchUut9.Busy;
   TraceOut_Done[120] := BenchUut9.Done;
   BenchCalls := BenchCalls + 1;
 121:
   BenchUut9.Start := FALSE;
   BenchUut9.Stop := FALSE;
   BenchUut9.Reset := FALSE;
   BenchUut9.ExtendDone := FALSE;
   BenchUut9.ClampDone := FALSE;
   BenchUut9.ReleaseDone := FALSE;
   BenchUut9.RetractDone := TRUE;
   TraceIn_Start[121] := BenchUut9.Start;
   TraceIn_Stop[121] := BenchUut9.Stop;
   TraceIn_Reset[121] := BenchUut9.Reset;
   TraceIn_ExtendDone[121] := BenchUut9.ExtendDone;
   TraceIn_ClampDone[121] := BenchUut9.ClampDone;
   TraceIn_ReleaseDone[121] := BenchUut9.ReleaseDone;
   TraceIn_RetractDone[121] := BenchUut9.RetractDone;
   BenchUut9();
   TraceOut_Extend[121] := BenchUut9.Extend;
   TraceOut_Clamp[121] := BenchUut9.Clamp;
   TraceOut_Release[121] := BenchUut9.Release;
   TraceOut_Retract[121] := BenchUut9.Retract;
   TraceOut_Busy[121] := BenchUut9.Busy;
   TraceOut_Done[121] := BenchUut9.Done;
   BenchCalls := BenchCalls + 1;
 122:
   BenchUut9.Start := TRUE;
   BenchUut9.Stop := FALSE;
   BenchUut9.Reset := FALSE;
   BenchUut9.ExtendDone := FALSE;
   BenchUut9.ClampDone := FALSE;
   BenchUut9.ReleaseDone := FALSE;
   BenchUut9.RetractDone := FALSE;
   TraceIn_Start[122] := BenchUut9.Start;
   TraceIn_Stop[122] := BenchUut9.Stop;
   TraceIn_Reset[122] := BenchUut9.Reset;
   TraceIn_ExtendDone[122] := BenchUut9.ExtendDone;
   TraceIn_ClampDone[122] := BenchUut9.ClampDone;
   TraceIn_ReleaseDone[122] := BenchUut9.ReleaseDone;
   TraceIn_RetractDone[122] := BenchUut9.RetractDone;
   BenchUut9();
   TraceOut_Extend[122] := BenchUut9.Extend;
   TraceOut_Clamp[122] := BenchUut9.Clamp;
   TraceOut_Release[122] := BenchUut9.Release;
   TraceOut_Retract[122] := BenchUut9.Retract;
   TraceOut_Busy[122] := BenchUut9.Busy;
   TraceOut_Done[122] := BenchUut9.Done;
   BenchCalls := BenchCalls + 1;
 123:
   BenchUut9.Start := FALSE;
   BenchUut9.Stop := FALSE;
   BenchUut9.Reset := TRUE;
   BenchUut9.ExtendDone := FALSE;
   BenchUut9.ClampDone := FALSE;
   BenchUut9.ReleaseDone := FALSE;
   BenchUut9.RetractDone := FALSE;
   TraceIn_Start[123] := BenchUut9.Start;
   TraceIn_Stop[123] := BenchUut9.Stop;
   TraceIn_Reset[123] := BenchUut9.Reset;
   TraceIn_ExtendDone[123] := BenchUut9.ExtendDone;
   TraceIn_ClampDone[123] := BenchUut9.ClampDone;
   TraceIn_ReleaseDone[123] := BenchUut9.ReleaseDone;
   TraceIn_RetractDone[123] := BenchUut9.RetractDone;
   BenchUut9();
   TraceOut_Extend[123] := BenchUut9.Extend;
   TraceOut_Clamp[123] := BenchUut9.Clamp;
   TraceOut_Release[123] := BenchUut9.Release;
   TraceOut_Retract[123] := BenchUut9.Retract;
   TraceOut_Busy[123] := BenchUut9.Busy;
   TraceOut_Done[123] := BenchUut9.Done;
   BenchCalls := BenchCalls + 1;
 124:
   BenchUut9.Start := FALSE;
   BenchUut9.Stop := FALSE;
   BenchUut9.Reset := TRUE;
   BenchUut9.ExtendDone := FALSE;
   BenchUut9.ClampDone := TRUE;
   BenchUut9.ReleaseDone := FALSE;
   BenchUut9.RetractDone := FALSE;
   TraceIn_Start[124] := BenchUut9.Start;
   TraceIn_Stop[124] := BenchUut9.Stop;
   TraceIn_Reset[124] := BenchUut9.Reset;
   TraceIn_ExtendDone[124] := BenchUut9.ExtendDone;
   TraceIn_ClampDone[124] := BenchUut9.ClampDone;
   TraceIn_ReleaseDone[124] := BenchUut9.ReleaseDone;
   TraceIn_RetractDone[124] := BenchUut9.RetractDone;
   BenchUut9();
   TraceOut_Extend[124] := BenchUut9.Extend;
   TraceOut_Clamp[124] := BenchUut9.Clamp;
   TraceOut_Release[124] := BenchUut9.Release;
   TraceOut_Retract[124] := BenchUut9.Retract;
   TraceOut_Busy[124] := BenchUut9.Busy;
   TraceOut_Done[124] := BenchUut9.Done;
   BenchCalls := BenchCalls + 1;
 125:
   BenchUut9.Start := FALSE;
   BenchUut9.Stop := FALSE;
   BenchUut9.Reset := TRUE;
   BenchUut9.ExtendDone := FALSE;
   BenchUut9.ClampDone := TRUE;
   BenchUut9.ReleaseDone := FALSE;
   BenchUut9.RetractDone := FALSE;
   TraceIn_Start[125] := BenchUut9.Start;
   TraceIn_Stop[125] := BenchUut9.Stop;
   TraceIn_Reset[125] := BenchUut9.Reset;
   TraceIn_ExtendDone[125] := BenchUut9.ExtendDone;
   TraceIn_ClampDone[125] := BenchUut9.ClampDone;
   TraceIn_ReleaseDone[125] := BenchUut9.ReleaseDone;
   TraceIn_RetractDone[125] := BenchUut9.RetractDone;
   BenchUut9();
   TraceOut_Extend[125] := BenchUut9.Extend;
   TraceOut_Clamp[125] := BenchUut9.Clamp;
   TraceOut_Release[125] := BenchUut9.Release;
   TraceOut_Retract[125] := BenchUut9.Retract;
   TraceOut_Busy[125] := BenchUut9.Busy;
   TraceOut_Done[125] := BenchUut9.Done;
   BenchCalls := BenchCalls + 1;
 126:
   BenchUut10.Start := TRUE;
   BenchUut10.Stop := FALSE;
   BenchUut10.Reset := FALSE;
   BenchUut10.ExtendDone := FALSE;
   BenchUut10.ClampDone := FALSE;
   BenchUut10.ReleaseDone := FALSE;
   BenchUut10.RetractDone := FALSE;
   TraceIn_Start[126] := BenchUut10.Start;
   TraceIn_Stop[126] := BenchUut10.Stop;
   TraceIn_Reset[126] := BenchUut10.Reset;
   TraceIn_ExtendDone[126] := BenchUut10.ExtendDone;
   TraceIn_ClampDone[126] := BenchUut10.ClampDone;
   TraceIn_ReleaseDone[126] := BenchUut10.ReleaseDone;
   TraceIn_RetractDone[126] := BenchUut10.RetractDone;
   BenchUut10();
   TraceOut_Extend[126] := BenchUut10.Extend;
   TraceOut_Clamp[126] := BenchUut10.Clamp;
   TraceOut_Release[126] := BenchUut10.Release;
   TraceOut_Retract[126] := BenchUut10.Retract;
   TraceOut_Busy[126] := BenchUut10.Busy;
   TraceOut_Done[126] := BenchUut10.Done;
   BenchCalls := BenchCalls + 1;
 127:
   BenchUut10.Start := TRUE;
   BenchUut10.Stop := FALSE;
   BenchUut10.Reset := FALSE;
   BenchUut10.ExtendDone := FALSE;
   BenchUut10.ClampDone := FALSE;
   BenchUut10.ReleaseDone := FALSE;
   BenchUut10.RetractDone := TRUE;
   TraceIn_Start[127] := BenchUut10.Start;
   TraceIn_Stop[127] := BenchUut10.Stop;
   TraceIn_Reset[127] := BenchUut10.Reset;
   TraceIn_ExtendDone[127] := BenchUut10.ExtendDone;
   TraceIn_ClampDone[127] := BenchUut10.ClampDone;
   TraceIn_ReleaseDone[127] := BenchUut10.ReleaseDone;
   TraceIn_RetractDone[127] := BenchUut10.RetractDone;
   BenchUut10();
   TraceOut_Extend[127] := BenchUut10.Extend;
   TraceOut_Clamp[127] := BenchUut10.Clamp;
   TraceOut_Release[127] := BenchUut10.Release;
   TraceOut_Retract[127] := BenchUut10.Retract;
   TraceOut_Busy[127] := BenchUut10.Busy;
   TraceOut_Done[127] := BenchUut10.Done;
   BenchCalls := BenchCalls + 1;
 128:
   BenchUut10.Start := FALSE;
   BenchUut10.Stop := FALSE;
   BenchUut10.Reset := FALSE;
   BenchUut10.ExtendDone := FALSE;
   BenchUut10.ClampDone := FALSE;
   BenchUut10.ReleaseDone := FALSE;
   BenchUut10.RetractDone := FALSE;
   TraceIn_Start[128] := BenchUut10.Start;
   TraceIn_Stop[128] := BenchUut10.Stop;
   TraceIn_Reset[128] := BenchUut10.Reset;
   TraceIn_ExtendDone[128] := BenchUut10.ExtendDone;
   TraceIn_ClampDone[128] := BenchUut10.ClampDone;
   TraceIn_ReleaseDone[128] := BenchUut10.ReleaseDone;
   TraceIn_RetractDone[128] := BenchUut10.RetractDone;
   BenchUut10();
   TraceOut_Extend[128] := BenchUut10.Extend;
   TraceOut_Clamp[128] := BenchUut10.Clamp;
   TraceOut_Release[128] := BenchUut10.Release;
   TraceOut_Retract[128] := BenchUut10.Retract;
   TraceOut_Busy[128] := BenchUut10.Busy;
   TraceOut_Done[128] := BenchUut10.Done;
   BenchCalls := BenchCalls + 1;
 129:
   BenchUut10.Start := FALSE;
   BenchUut10.Stop := FALSE;
   BenchUut10.Reset := FALSE;
   BenchUut10.ExtendDone := TRUE;
   BenchUut10.ClampDone := FALSE;
   BenchUut10.ReleaseDone := FALSE;
   BenchUut10.RetractDone := FALSE;
   TraceIn_Start[129] := BenchUut10.Start;
   TraceIn_Stop[129] := BenchUut10.Stop;
   TraceIn_Reset[129] := BenchUut10.Reset;
   TraceIn_ExtendDone[129] := BenchUut10.ExtendDone;
   TraceIn_ClampDone[129] := BenchUut10.ClampDone;
   TraceIn_ReleaseDone[129] := BenchUut10.ReleaseDone;
   TraceIn_RetractDone[129] := BenchUut10.RetractDone;
   BenchUut10();
   TraceOut_Extend[129] := BenchUut10.Extend;
   TraceOut_Clamp[129] := BenchUut10.Clamp;
   TraceOut_Release[129] := BenchUut10.Release;
   TraceOut_Retract[129] := BenchUut10.Retract;
   TraceOut_Busy[129] := BenchUut10.Busy;
   TraceOut_Done[129] := BenchUut10.Done;
   BenchCalls := BenchCalls + 1;
 130:
   BenchUut10.Start := FALSE;
   BenchUut10.Stop := FALSE;
   BenchUut10.Reset := FALSE;
   BenchUut10.ExtendDone := FALSE;
   BenchUut10.ClampDone := TRUE;
   BenchUut10.ReleaseDone := FALSE;
   BenchUut10.RetractDone := FALSE;
   TraceIn_Start[130] := BenchUut10.Start;
   TraceIn_Stop[130] := BenchUut10.Stop;
   TraceIn_Reset[130] := BenchUut10.Reset;
   TraceIn_ExtendDone[130] := BenchUut10.ExtendDone;
   TraceIn_ClampDone[130] := BenchUut10.ClampDone;
   TraceIn_ReleaseDone[130] := BenchUut10.ReleaseDone;
   TraceIn_RetractDone[130] := BenchUut10.RetractDone;
   BenchUut10();
   TraceOut_Extend[130] := BenchUut10.Extend;
   TraceOut_Clamp[130] := BenchUut10.Clamp;
   TraceOut_Release[130] := BenchUut10.Release;
   TraceOut_Retract[130] := BenchUut10.Retract;
   TraceOut_Busy[130] := BenchUut10.Busy;
   TraceOut_Done[130] := BenchUut10.Done;
   BenchCalls := BenchCalls + 1;
 131:
   BenchUut10.Start := FALSE;
   BenchUut10.Stop := FALSE;
   BenchUut10.Reset := FALSE;
   BenchUut10.ExtendDone := FALSE;
   BenchUut10.ClampDone := FALSE;
   BenchUut10.ReleaseDone := TRUE;
   BenchUut10.RetractDone := FALSE;
   TraceIn_Start[131] := BenchUut10.Start;
   TraceIn_Stop[131] := BenchUut10.Stop;
   TraceIn_Reset[131] := BenchUut10.Reset;
   TraceIn_ExtendDone[131] := BenchUut10.ExtendDone;
   TraceIn_ClampDone[131] := BenchUut10.ClampDone;
   TraceIn_ReleaseDone[131] := BenchUut10.ReleaseDone;
   TraceIn_RetractDone[131] := BenchUut10.RetractDone;
   BenchUut10();
   TraceOut_Extend[131] := BenchUut10.Extend;
   TraceOut_Clamp[131] := BenchUut10.Clamp;
   TraceOut_Release[131] := BenchUut10.Release;
   TraceOut_Retract[131] := BenchUut10.Retract;
   TraceOut_Busy[131] := BenchUut10.Busy;
   TraceOut_Done[131] := BenchUut10.Done;
   BenchCalls := BenchCalls + 1;
 132:
   BenchUut10.Start := FALSE;
   BenchUut10.Stop := FALSE;
   BenchUut10.Reset := FALSE;
   BenchUut10.ExtendDone := FALSE;
   BenchUut10.ClampDone := FALSE;
   BenchUut10.ReleaseDone := FALSE;
   BenchUut10.RetractDone := TRUE;
   TraceIn_Start[132] := BenchUut10.Start;
   TraceIn_Stop[132] := BenchUut10.Stop;
   TraceIn_Reset[132] := BenchUut10.Reset;
   TraceIn_ExtendDone[132] := BenchUut10.ExtendDone;
   TraceIn_ClampDone[132] := BenchUut10.ClampDone;
   TraceIn_ReleaseDone[132] := BenchUut10.ReleaseDone;
   TraceIn_RetractDone[132] := BenchUut10.RetractDone;
   BenchUut10();
   TraceOut_Extend[132] := BenchUut10.Extend;
   TraceOut_Clamp[132] := BenchUut10.Clamp;
   TraceOut_Release[132] := BenchUut10.Release;
   TraceOut_Retract[132] := BenchUut10.Retract;
   TraceOut_Busy[132] := BenchUut10.Busy;
   TraceOut_Done[132] := BenchUut10.Done;
   BenchCalls := BenchCalls + 1;
 133:
   BenchUut10.Start := TRUE;
   BenchUut10.Stop := FALSE;
   BenchUut10.Reset := FALSE;
   BenchUut10.ExtendDone := FALSE;
   BenchUut10.ClampDone := FALSE;
   BenchUut10.ReleaseDone := FALSE;
   BenchUut10.RetractDone := FALSE;
   TraceIn_Start[133] := BenchUut10.Start;
   TraceIn_Stop[133] := BenchUut10.Stop;
   TraceIn_Reset[133] := BenchUut10.Reset;
   TraceIn_ExtendDone[133] := BenchUut10.ExtendDone;
   TraceIn_ClampDone[133] := BenchUut10.ClampDone;
   TraceIn_ReleaseDone[133] := BenchUut10.ReleaseDone;
   TraceIn_RetractDone[133] := BenchUut10.RetractDone;
   BenchUut10();
   TraceOut_Extend[133] := BenchUut10.Extend;
   TraceOut_Clamp[133] := BenchUut10.Clamp;
   TraceOut_Release[133] := BenchUut10.Release;
   TraceOut_Retract[133] := BenchUut10.Retract;
   TraceOut_Busy[133] := BenchUut10.Busy;
   TraceOut_Done[133] := BenchUut10.Done;
   BenchCalls := BenchCalls + 1;
 134:
   BenchUut10.Start := FALSE;
   BenchUut10.Stop := FALSE;
   BenchUut10.Reset := TRUE;
   BenchUut10.ExtendDone := FALSE;
   BenchUut10.ClampDone := FALSE;
   BenchUut10.ReleaseDone := FALSE;
   BenchUut10.RetractDone := FALSE;
   TraceIn_Start[134] := BenchUut10.Start;
   TraceIn_Stop[134] := BenchUut10.Stop;
   TraceIn_Reset[134] := BenchUut10.Reset;
   TraceIn_ExtendDone[134] := BenchUut10.ExtendDone;
   TraceIn_ClampDone[134] := BenchUut10.ClampDone;
   TraceIn_ReleaseDone[134] := BenchUut10.ReleaseDone;
   TraceIn_RetractDone[134] := BenchUut10.RetractDone;
   BenchUut10();
   TraceOut_Extend[134] := BenchUut10.Extend;
   TraceOut_Clamp[134] := BenchUut10.Clamp;
   TraceOut_Release[134] := BenchUut10.Release;
   TraceOut_Retract[134] := BenchUut10.Retract;
   TraceOut_Busy[134] := BenchUut10.Busy;
   TraceOut_Done[134] := BenchUut10.Done;
   BenchCalls := BenchCalls + 1;
 135:
   BenchUut10.Start := FALSE;
   BenchUut10.Stop := FALSE;
   BenchUut10.Reset := TRUE;
   BenchUut10.ExtendDone := FALSE;
   BenchUut10.ClampDone := FALSE;
   BenchUut10.ReleaseDone := TRUE;
   BenchUut10.RetractDone := FALSE;
   TraceIn_Start[135] := BenchUut10.Start;
   TraceIn_Stop[135] := BenchUut10.Stop;
   TraceIn_Reset[135] := BenchUut10.Reset;
   TraceIn_ExtendDone[135] := BenchUut10.ExtendDone;
   TraceIn_ClampDone[135] := BenchUut10.ClampDone;
   TraceIn_ReleaseDone[135] := BenchUut10.ReleaseDone;
   TraceIn_RetractDone[135] := BenchUut10.RetractDone;
   BenchUut10();
   TraceOut_Extend[135] := BenchUut10.Extend;
   TraceOut_Clamp[135] := BenchUut10.Clamp;
   TraceOut_Release[135] := BenchUut10.Release;
   TraceOut_Retract[135] := BenchUut10.Retract;
   TraceOut_Busy[135] := BenchUut10.Busy;
   TraceOut_Done[135] := BenchUut10.Done;
   BenchCalls := BenchCalls + 1;
 136:
   BenchUut10.Start := FALSE;
   BenchUut10.Stop := FALSE;
   BenchUut10.Reset := TRUE;
   BenchUut10.ExtendDone := FALSE;
   BenchUut10.ClampDone := FALSE;
   BenchUut10.ReleaseDone := TRUE;
   BenchUut10.RetractDone := FALSE;
   TraceIn_Start[136] := BenchUut10.Start;
   TraceIn_Stop[136] := BenchUut10.Stop;
   TraceIn_Reset[136] := BenchUut10.Reset;
   TraceIn_ExtendDone[136] := BenchUut10.ExtendDone;
   TraceIn_ClampDone[136] := BenchUut10.ClampDone;
   TraceIn_ReleaseDone[136] := BenchUut10.ReleaseDone;
   TraceIn_RetractDone[136] := BenchUut10.RetractDone;
   BenchUut10();
   TraceOut_Extend[136] := BenchUut10.Extend;
   TraceOut_Clamp[136] := BenchUut10.Clamp;
   TraceOut_Release[136] := BenchUut10.Release;
   TraceOut_Retract[136] := BenchUut10.Retract;
   TraceOut_Busy[136] := BenchUut10.Busy;
   TraceOut_Done[136] := BenchUut10.Done;
   BenchCalls := BenchCalls + 1;
 137:
   BenchUut11.Start := TRUE;
   BenchUut11.Stop := FALSE;
   BenchUut11.Reset := FALSE;
   BenchUut11.ExtendDone := FALSE;
   BenchUut11.ClampDone := FALSE;
   BenchUut11.ReleaseDone := FALSE;
   BenchUut11.RetractDone := FALSE;
   TraceIn_Start[137] := BenchUut11.Start;
   TraceIn_Stop[137] := BenchUut11.Stop;
   TraceIn_Reset[137] := BenchUut11.Reset;
   TraceIn_ExtendDone[137] := BenchUut11.ExtendDone;
   TraceIn_ClampDone[137] := BenchUut11.ClampDone;
   TraceIn_ReleaseDone[137] := BenchUut11.ReleaseDone;
   TraceIn_RetractDone[137] := BenchUut11.RetractDone;
   BenchUut11();
   TraceOut_Extend[137] := BenchUut11.Extend;
   TraceOut_Clamp[137] := BenchUut11.Clamp;
   TraceOut_Release[137] := BenchUut11.Release;
   TraceOut_Retract[137] := BenchUut11.Retract;
   TraceOut_Busy[137] := BenchUut11.Busy;
   TraceOut_Done[137] := BenchUut11.Done;
   BenchCalls := BenchCalls + 1;
 138:
   BenchUut11.Start := TRUE;
   BenchUut11.Stop := FALSE;
   BenchUut11.Reset := FALSE;
   BenchUut11.ExtendDone := FALSE;
   BenchUut11.ClampDone := FALSE;
   BenchUut11.ReleaseDone := FALSE;
   BenchUut11.RetractDone := TRUE;
   TraceIn_Start[138] := BenchUut11.Start;
   TraceIn_Stop[138] := BenchUut11.Stop;
   TraceIn_Reset[138] := BenchUut11.Reset;
   TraceIn_ExtendDone[138] := BenchUut11.ExtendDone;
   TraceIn_ClampDone[138] := BenchUut11.ClampDone;
   TraceIn_ReleaseDone[138] := BenchUut11.ReleaseDone;
   TraceIn_RetractDone[138] := BenchUut11.RetractDone;
   BenchUut11();
   TraceOut_Extend[138] := BenchUut11.Extend;
   TraceOut_Clamp[138] := BenchUut11.Clamp;
   TraceOut_Release[138] := BenchUut11.Release;
   TraceOut_Retract[138] := BenchUut11.Retract;
   TraceOut_Busy[138] := BenchUut11.Busy;
   TraceOut_Done[138] := BenchUut11.Done;
   BenchCalls := BenchCalls + 1;
 139:
   BenchUut11.Start := FALSE;
   BenchUut11.Stop := FALSE;
   BenchUut11.Reset := FALSE;
   BenchUut11.ExtendDone := FALSE;
   BenchUut11.ClampDone := FALSE;
   BenchUut11.ReleaseDone := FALSE;
   BenchUut11.RetractDone := FALSE;
   TraceIn_Start[139] := BenchUut11.Start;
   TraceIn_Stop[139] := BenchUut11.Stop;
   TraceIn_Reset[139] := BenchUut11.Reset;
   TraceIn_ExtendDone[139] := BenchUut11.ExtendDone;
   TraceIn_ClampDone[139] := BenchUut11.ClampDone;
   TraceIn_ReleaseDone[139] := BenchUut11.ReleaseDone;
   TraceIn_RetractDone[139] := BenchUut11.RetractDone;
   BenchUut11();
   TraceOut_Extend[139] := BenchUut11.Extend;
   TraceOut_Clamp[139] := BenchUut11.Clamp;
   TraceOut_Release[139] := BenchUut11.Release;
   TraceOut_Retract[139] := BenchUut11.Retract;
   TraceOut_Busy[139] := BenchUut11.Busy;
   TraceOut_Done[139] := BenchUut11.Done;
   BenchCalls := BenchCalls + 1;
 140:
   BenchUut11.Start := FALSE;
   BenchUut11.Stop := FALSE;
   BenchUut11.Reset := FALSE;
   BenchUut11.ExtendDone := TRUE;
   BenchUut11.ClampDone := FALSE;
   BenchUut11.ReleaseDone := FALSE;
   BenchUut11.RetractDone := FALSE;
   TraceIn_Start[140] := BenchUut11.Start;
   TraceIn_Stop[140] := BenchUut11.Stop;
   TraceIn_Reset[140] := BenchUut11.Reset;
   TraceIn_ExtendDone[140] := BenchUut11.ExtendDone;
   TraceIn_ClampDone[140] := BenchUut11.ClampDone;
   TraceIn_ReleaseDone[140] := BenchUut11.ReleaseDone;
   TraceIn_RetractDone[140] := BenchUut11.RetractDone;
   BenchUut11();
   TraceOut_Extend[140] := BenchUut11.Extend;
   TraceOut_Clamp[140] := BenchUut11.Clamp;
   TraceOut_Release[140] := BenchUut11.Release;
   TraceOut_Retract[140] := BenchUut11.Retract;
   TraceOut_Busy[140] := BenchUut11.Busy;
   TraceOut_Done[140] := BenchUut11.Done;
   BenchCalls := BenchCalls + 1;
 141:
   BenchUut11.Start := FALSE;
   BenchUut11.Stop := FALSE;
   BenchUut11.Reset := FALSE;
   BenchUut11.ExtendDone := FALSE;
   BenchUut11.ClampDone := TRUE;
   BenchUut11.ReleaseDone := FALSE;
   BenchUut11.RetractDone := FALSE;
   TraceIn_Start[141] := BenchUut11.Start;
   TraceIn_Stop[141] := BenchUut11.Stop;
   TraceIn_Reset[141] := BenchUut11.Reset;
   TraceIn_ExtendDone[141] := BenchUut11.ExtendDone;
   TraceIn_ClampDone[141] := BenchUut11.ClampDone;
   TraceIn_ReleaseDone[141] := BenchUut11.ReleaseDone;
   TraceIn_RetractDone[141] := BenchUut11.RetractDone;
   BenchUut11();
   TraceOut_Extend[141] := BenchUut11.Extend;
   TraceOut_Clamp[141] := BenchUut11.Clamp;
   TraceOut_Release[141] := BenchUut11.Release;
   TraceOut_Retract[141] := BenchUut11.Retract;
   TraceOut_Busy[141] := BenchUut11.Busy;
   TraceOut_Done[141] := BenchUut11.Done;
   BenchCalls := BenchCalls + 1;
 142:
   BenchUut11.Start := FALSE;
   BenchUut11.Stop := FALSE;
   BenchUut11.Reset := FALSE;
   BenchUut11.ExtendDone := FALSE;
   BenchUut11.ClampDone := FALSE;
   BenchUut11.ReleaseDone := TRUE;
   BenchUut11.RetractDone := FALSE;
   TraceIn_Start[142] := BenchUut11.Start;
   TraceIn_Stop[142] := BenchUut11.Stop;
   TraceIn_Reset[142] := BenchUut11.Reset;
   TraceIn_ExtendDone[142] := BenchUut11.ExtendDone;
   TraceIn_ClampDone[142] := BenchUut11.ClampDone;
   TraceIn_ReleaseDone[142] := BenchUut11.ReleaseDone;
   TraceIn_RetractDone[142] := BenchUut11.RetractDone;
   BenchUut11();
   TraceOut_Extend[142] := BenchUut11.Extend;
   TraceOut_Clamp[142] := BenchUut11.Clamp;
   TraceOut_Release[142] := BenchUut11.Release;
   TraceOut_Retract[142] := BenchUut11.Retract;
   TraceOut_Busy[142] := BenchUut11.Busy;
   TraceOut_Done[142] := BenchUut11.Done;
   BenchCalls := BenchCalls + 1;
 143:
   BenchUut11.Start := FALSE;
   BenchUut11.Stop := FALSE;
   BenchUut11.Reset := FALSE;
   BenchUut11.ExtendDone := FALSE;
   BenchUut11.ClampDone := FALSE;
   BenchUut11.ReleaseDone := FALSE;
   BenchUut11.RetractDone := TRUE;
   TraceIn_Start[143] := BenchUut11.Start;
   TraceIn_Stop[143] := BenchUut11.Stop;
   TraceIn_Reset[143] := BenchUut11.Reset;
   TraceIn_ExtendDone[143] := BenchUut11.ExtendDone;
   TraceIn_ClampDone[143] := BenchUut11.ClampDone;
   TraceIn_ReleaseDone[143] := BenchUut11.ReleaseDone;
   TraceIn_RetractDone[143] := BenchUut11.RetractDone;
   BenchUut11();
   TraceOut_Extend[143] := BenchUut11.Extend;
   TraceOut_Clamp[143] := BenchUut11.Clamp;
   TraceOut_Release[143] := BenchUut11.Release;
   TraceOut_Retract[143] := BenchUut11.Retract;
   TraceOut_Busy[143] := BenchUut11.Busy;
   TraceOut_Done[143] := BenchUut11.Done;
   BenchCalls := BenchCalls + 1;
 144:
   BenchUut11.Start := TRUE;
   BenchUut11.Stop := FALSE;
   BenchUut11.Reset := FALSE;
   BenchUut11.ExtendDone := FALSE;
   BenchUut11.ClampDone := FALSE;
   BenchUut11.ReleaseDone := FALSE;
   BenchUut11.RetractDone := FALSE;
   TraceIn_Start[144] := BenchUut11.Start;
   TraceIn_Stop[144] := BenchUut11.Stop;
   TraceIn_Reset[144] := BenchUut11.Reset;
   TraceIn_ExtendDone[144] := BenchUut11.ExtendDone;
   TraceIn_ClampDone[144] := BenchUut11.ClampDone;
   TraceIn_ReleaseDone[144] := BenchUut11.ReleaseDone;
   TraceIn_RetractDone[144] := BenchUut11.RetractDone;
   BenchUut11();
   TraceOut_Extend[144] := BenchUut11.Extend;
   TraceOut_Clamp[144] := BenchUut11.Clamp;
   TraceOut_Release[144] := BenchUut11.Release;
   TraceOut_Retract[144] := BenchUut11.Retract;
   TraceOut_Busy[144] := BenchUut11.Busy;
   TraceOut_Done[144] := BenchUut11.Done;
   BenchCalls := BenchCalls + 1;
 145:
   BenchUut11.Start := FALSE;
   BenchUut11.Stop := FALSE;
   BenchUut11.Reset := TRUE;
   BenchUut11.ExtendDone := FALSE;
   BenchUut11.ClampDone := FALSE;
   BenchUut11.ReleaseDone := FALSE;
   BenchUut11.RetractDone := FALSE;
   TraceIn_Start[145] := BenchUut11.Start;
   TraceIn_Stop[145] := BenchUut11.Stop;
   TraceIn_Reset[145] := BenchUut11.Reset;
   TraceIn_ExtendDone[145] := BenchUut11.ExtendDone;
   TraceIn_ClampDone[145] := BenchUut11.ClampDone;
   TraceIn_ReleaseDone[145] := BenchUut11.ReleaseDone;
   TraceIn_RetractDone[145] := BenchUut11.RetractDone;
   BenchUut11();
   TraceOut_Extend[145] := BenchUut11.Extend;
   TraceOut_Clamp[145] := BenchUut11.Clamp;
   TraceOut_Release[145] := BenchUut11.Release;
   TraceOut_Retract[145] := BenchUut11.Retract;
   TraceOut_Busy[145] := BenchUut11.Busy;
   TraceOut_Done[145] := BenchUut11.Done;
   BenchCalls := BenchCalls + 1;
 146:
   BenchUut11.Start := FALSE;
   BenchUut11.Stop := FALSE;
   BenchUut11.Reset := TRUE;
   BenchUut11.ExtendDone := FALSE;
   BenchUut11.ClampDone := FALSE;
   BenchUut11.ReleaseDone := FALSE;
   BenchUut11.RetractDone := TRUE;
   TraceIn_Start[146] := BenchUut11.Start;
   TraceIn_Stop[146] := BenchUut11.Stop;
   TraceIn_Reset[146] := BenchUut11.Reset;
   TraceIn_ExtendDone[146] := BenchUut11.ExtendDone;
   TraceIn_ClampDone[146] := BenchUut11.ClampDone;
   TraceIn_ReleaseDone[146] := BenchUut11.ReleaseDone;
   TraceIn_RetractDone[146] := BenchUut11.RetractDone;
   BenchUut11();
   TraceOut_Extend[146] := BenchUut11.Extend;
   TraceOut_Clamp[146] := BenchUut11.Clamp;
   TraceOut_Release[146] := BenchUut11.Release;
   TraceOut_Retract[146] := BenchUut11.Retract;
   TraceOut_Busy[146] := BenchUut11.Busy;
   TraceOut_Done[146] := BenchUut11.Done;
   BenchCalls := BenchCalls + 1;
 147:
   BenchUut11.Start := FALSE;
   BenchUut11.Stop := FALSE;
   BenchUut11.Reset := TRUE;
   BenchUut11.ExtendDone := FALSE;
   BenchUut11.ClampDone := FALSE;
   BenchUut11.ReleaseDone := FALSE;
   BenchUut11.RetractDone := TRUE;
   TraceIn_Start[147] := BenchUut11.Start;
   TraceIn_Stop[147] := BenchUut11.Stop;
   TraceIn_Reset[147] := BenchUut11.Reset;
   TraceIn_ExtendDone[147] := BenchUut11.ExtendDone;
   TraceIn_ClampDone[147] := BenchUut11.ClampDone;
   TraceIn_ReleaseDone[147] := BenchUut11.ReleaseDone;
   TraceIn_RetractDone[147] := BenchUut11.RetractDone;
   BenchUut11();
   TraceOut_Extend[147] := BenchUut11.Extend;
   TraceOut_Clamp[147] := BenchUut11.Clamp;
   TraceOut_Release[147] := BenchUut11.Release;
   TraceOut_Retract[147] := BenchUut11.Retract;
   TraceOut_Busy[147] := BenchUut11.Busy;
   TraceOut_Done[147] := BenchUut11.Done;
   BenchCalls := BenchCalls + 1;
 END_CASE;
 BenchStep := BenchStep + 1;
 IF BenchStep >= 148 THEN BenchDone := TRUE; END_IF;
END_IF;
END_PROGRAM
